NETWORK
TITLE = Station Sicher Pos3.0
      AN    "POS3_0_Prodiag_DB".State.C1;

      =     "HMI_BETR_ART_POS".POS3_0.Status_Sicher;

END_FUNCTION_BLOCK

FUNCTION_BLOCK "Melden_VisuAllgemein"   // FB127, LAD
{ S7_Optimized_Access := 'TRUE' }
// stored: MemoryReserve 100, SetENOAutomatically false
   VAR
      Register_leer : "Teile Status";
      auf_Seite_Richten { S7_SetPoint := 'True'} : Bool;
      Flanke_Bildwechsel { S7_SetPoint := 'True'} : R_TRIG;
      Bild_tmp { S7_SetPoint := 'True'} : DInt;
      WartezeitSicherung_Reset { S7_SetPoint := 'True'} : TON_TIME;
      Flanke_Türe8_schließen { S7_SetPoint := 'True'} : R_TRIG;
      Flanke_Türe8_öffnen { S7_SetPoint := 'True'} : R_TRIG;
   END_VAR
   VAR RETAIN
      Artikelnummer_tmp { ExternalAccessible := 'False'; ExternalVisible := 'False'; ExternalWritable := 'False'} : String;
   END_VAR
   VAR
      VZ_Leerfahren { S7_SetPoint := 'True'} : TON_TIME;
   END_VAR
   VAR_TEMP
      test : Bool;
   END_VAR
BEGIN

REGION Network 1 (SCL): Richten oder Einzelschrittseite aufgerufen
   CASE "HMI_SYS"."Aktueller Bildschirm" OF
       75:
           #auf_Seite_Richten := true;
       ELSE
           #auf_Seite_Richten := false;
   END_CASE;
END_REGION

REGION Network 2 (SCL): Artikel wurde gewechselt


   IF #Artikelnummer_tmp <> "HMI_COM".Artikelnummer_String THEN
       "HMI_COM".Artikel_gewechselt := true;
       #Artikelnummer_tmp := "HMI_COM".Artikelnummer_String;
   ELSIF "HMI_COM".Grundstellung_Gesamt AND  "HMI_COM".Artikel_gewechselt THEN

       "HMI_COM".Artikel_gewechselt := false;

   END_IF;
END_REGION

NETWORK
TITLE = Übergabe Anwahl Richten
      A     #auf_Seite_Richten;
      JC    m003;

      JU    m001;
m003: NOP   0;

      A     "03_Betriebsart_DB"."NOT-HALT OK";
      A     "03_Betriebsart_DB"."Schutztüren OK";
      JCN   m001;


      A     "HMI_COM".Richten_Gesamtanlage;
      JCN   m002;

      SET;
      S     "HMI_BETR_ART_POS".POS3_0.Taster_Anwahl_GS;


m002: NOP   0;

      A     "HMI_BETR_ART_POS".POS3_0.Taster_Anwahl_GS;
      S     "POS3_0_Signal".Station.SK_Freigabe_Richten;
      =     "POS3_0_Signal".Schrittkette.INIT_SQ;
      R     "HMI_BETR_ART_POS".POS3_0.Taster_Anwahl_GS;


      A     "HMI_COM".Richten_Gesamtanlage;
      R     "HMI_COM".Richten_Gesamtanlage;

m001: NOP   0;


NETWORK
TITLE = Tippbetrieb Aktiv
      A     "POS3_0_Signal".Schrittkette.AUTO_ON;


      =     "HMI_COM".Einzelschritt.Status_Anw;


NETWORK
TITLE = Antriebe sind Ein
      SET;

      =     "HMI_COM".Antriebe_sind_EIN;

REGION Network 6 (SCL): Übergabe Türen Not Halt
   // Allgemeine HMI Übergabe 

   "HMI_COM"."NOT-HALT_OK" := "03_Betriebsart_DB"."NOT-HALT OK";
   "HMI_COM".TUERE_OK := "03_Betriebsart_DB"."Schutztüren OK";




   // Übergabe welche Tür ist nicht verriegelt
   REGION Türen


       "HMI_COM".Tür_offen[1] := "DE_Rueckfuehrung_Tuer_1" AND ("03_Betriebsart_DB".BA_Automatik OR "03_Betriebsart_DB".BA_Manuell OR "03_Betriebsart_DB".BA_Richten);
       "HMI_COM".Tür_offen[2] := "DE_Rueckfuehrung_Tuer_2" AND ("03_Betriebsart_DB".BA_Automatik OR "03_Betriebsart_DB".BA_Manuell OR "03_Betriebsart_DB".BA_Richten);
    //   "HMI_COM".Tür_offen[3] := "DE_Rueckfuehrung_Tuer_3" AND ("03_Betriebsart_DB".BA_Automatik OR "03_Betriebsart_DB".BA_Manuell OR "03_Betriebsart_DB".BA_Richten);
    //   "HMI_COM".Tür_offen[4] := "DE_Rueckfuehrung_Tuer_4" AND ("03_Betriebsart_DB".BA_Automatik OR "03_Betriebsart_DB".BA_Manuell OR "03_Betriebsart_DB".BA_Richten);
    //   "HMI_COM".Tür_offen[5] := "DE_Rueckfuehrung_Tuer_5" AND ("03_Betriebsart_DB".BA_Automatik OR "03_Betriebsart_DB".BA_Manuell OR "03_Betriebsart_DB".BA_Richten);
    //   "HMI_COM".Tür_offen[6] := "DE_Rueckfuehrung_Tuer_6" AND ("03_Betriebsart_DB".BA_Automatik OR "03_Betriebsart_DB".BA_Manuell OR "03_Betriebsart_DB".BA_Richten);
    //   "HMI_COM".Tür_offen[7] := "DE2_0_Rückführung Tür 7" AND ("03_Betriebsart_DB".BA_Automatik OR "03_Betriebsart_DB".BA_Manuell OR "03_Betriebsart_DB".BA_Richten);
    //   "HMI_COM".Tür_offen[8] := "DE2_1_Rückführung Tür 8" AND ("03_Betriebsart_DB".BA_Automatik OR "03_Betriebsart_DB".BA_Manuell OR "03_Betriebsart_DB".BA_Richten);
    (*   "HMI_COM".Tür_offen[9] := "DE2_1_Rückführung Tür 8" AND ("03_Betriebsart_DB".BA_Automatik OR "03_Betriebsart_DB".BA_Manuell OR "03_Betriebsart_DB".BA_Richten);
       "HMI_COM".Tür_offen[10] := "DE2_1_Rückführung Tür 8" AND ("03_Betriebsart_DB".BA_Automatik OR "03_Betriebsart_DB".BA_Manuell OR "03_Betriebsart_DB".BA_Richten);
       "HMI_COM".Tür_offen[11] := "DE2_1_Rückführung Tür 8" AND ("03_Betriebsart_DB".BA_Automatik OR "03_Betriebsart_DB".BA_Manuell OR "03_Betriebsart_DB".BA_Richten);
       "HMI_COM".Tür_offen[12] := "DE2_1_Rückführung Tür 8" AND ("03_Betriebsart_DB".BA_Automatik OR "03_Betriebsart_DB".BA_Manuell OR "03_Betriebsart_DB".BA_Richten);
       "HMI_COM".Tür_offen[13] := "DE2_1_Rückführung Tür 8" AND ("03_Betriebsart_DB".BA_Automatik OR "03_Betriebsart_DB".BA_Manuell OR "03_Betriebsart_DB".BA_Richten);
       "HMI_COM".Tür_offen[14] := "DE2_1_Rückführung Tür 8" AND ("03_Betriebsart_DB".BA_Automatik OR "03_Betriebsart_DB".BA_Manuell OR "03_Betriebsart_DB".BA_Richten);
       "HMI_COM".Tür_offen[15] := "DE2_1_Rückführung Tür 8" AND ("03_Betriebsart_DB".BA_Automatik OR "03_Betriebsart_DB".BA_Manuell OR "03_Betriebsart_DB".BA_Richten); *)
    //   "HMI_COM".Tür_offen[16] := "DE2_1_Rückführung Tür 8" AND ("03_Betriebsart_DB".BA_Automatik OR "03_Betriebsart_DB".BA_Manuell OR "03_Betriebsart_DB".BA_Richten);

   END_REGION
END_REGION

REGION Network 7 (SCL): Rücksetzen der Stationen bei Grundbild



   #Flanke_Bildwechsel(CLK:="03_Betriebsart_DB".BA_Manuell AND #Bild_tmp <> "HMI_SYS"."Aktueller Bildschirm" );



   IF #Flanke_Bildwechsel.Q THEN

       #Bild_tmp := "HMI_SYS"."Aktueller Bildschirm";

    //IF ("HMI_SYS"."Aktueller Bildschirm" = 10125) OR ("03_Betriebsart_DB"."NOT-HALT OK" = false) THEN

       "HMI_COM".Manuell_Zylinder1.Status := 0;
       "HMI_COM".Manuell_Zylinder2.Status := 0;
       "HMI_COM".Manuell_Zylinder3.Status := 0;
       "HMI_COM".Manuell_Zylinder4.Status := 0;

       "HMI_COM".Manuell_Zylinder1.GS := FALSE;
       "HMI_COM".Manuell_Zylinder1.AS1 := FALSE;
       "HMI_COM".Manuell_Zylinder2.GS := FALSE;
       "HMI_COM".Manuell_Zylinder2.AS1 := FALSE;
       "HMI_COM".Manuell_Zylinder3.GS := FALSE;
       "HMI_COM".Manuell_Zylinder3.AS1 := FALSE;
       "HMI_COM".Manuell_Zylinder4.GS := FALSE;
       "HMI_COM".Manuell_Zylinder4.AS1 := FALSE;

      "HMI_COM".Manuell_Zylinder1.DA_GS := FALSE;
       "HMI_COM".Manuell_Zylinder1.DA_AS1 := FALSE;
       "HMI_COM".Manuell_Zylinder2.DA_GS := FALSE;
       "HMI_COM".Manuell_Zylinder2.DA_AS1 := FALSE;
       "HMI_COM".Manuell_Zylinder3.DA_GS := FALSE;
       "HMI_COM".Manuell_Zylinder3.DA_AS1 := FALSE;
       "HMI_COM".Manuell_Zylinder4.DA_GS := FALSE;
       "HMI_COM".Manuell_Zylinder4.DA_AS1 := FALSE;
     END_IF;
END_REGION

REGION Network 8 (SCL): Übertragung und Verwaltung Register



   "HMI_COM".Speichern_Register := false;
END_REGION

REGION Network 9 (SCL): Rucksetzen wenn Register nicht gelöscht
   IF (("HMI_SYS"."Aktueller Bildschirm" = 10001) OR ("HMI_SYS"."Aktueller Bildschirm" = 10010) OR ("HMI_SYS"."Aktueller Bildschirm" = 10020)
       OR ("HMI_SYS"."Aktueller Bildschirm" = 10030)) THEN

       "HMI_BETR_ART_POS".POS3_0.Taster_Reset_Teilestatus := FALSE;
       "HMI_BETR_ART_POS".POS3_1.Taster_Reset_Teilestatus := FALSE;
       "HMI_BETR_ART_POS".POS3_2.Taster_Reset_Teilestatus := FALSE;
       "HMI_BETR_ART_POS".POS3_3.Taster_Reset_Teilestatus := FALSE;
       "HMI_BETR_ART_POS".POS3_4.Taster_Reset_Teilestatus := FALSE;
       "HMI_BETR_ART_POS".POS4_0_Zuführung.Taster_Reset_Teilestatus := FALSE;
       "HMI_BETR_ART_POS".POS5_0_Zuführung.Taster_Reset_Teilestatus := FALSE;
       "HMI_BETR_ART_POS".POS5_0.Taster_Reset_Teilestatus := FALSE;
       "HMI_BETR_ART_POS".POS6_0.Taster_Reset_Teilestatus := FALSE;
       "HMI_BETR_ART_POS".POS7_0.Taster_Reset_Teilestatus := FALSE;
       "HMI_BETR_ART_POS".POS7_1.Taster_Reset_Teilestatus := FALSE;
       "HMI_BETR_ART_POS".POS7_2.Taster_Reset_Teilestatus := FALSE;
       "HMI_BETR_ART_POS".POS7_3.Taster_Reset_Teilestatus := FALSE;
       "HMI_BETR_ART_POS".POS7_4.Taster_Reset_Teilestatus := FALSE;
       "HMI_BETR_ART_POS".POS8_0.Taster_Reset_Teilestatus := FALSE;
       "HMI_BETR_ART_POS".POS9_0.Taster_Reset_Teilestatus := FALSE;
       "HMI_BETR_ART_POS".POS9_1.Taster_Reset_Teilestatus := FALSE;
       "HMI_BETR_ART_POS".POS9_2.Taster_Reset_Teilestatus := FALSE;
       "HMI_BETR_ART_POS".POS9_3.Taster_Reset_Teilestatus := FALSE;
       "HMI_BETR_ART_POS".POS9_4.Taster_Reset_Teilestatus := FALSE;
       "HMI_BETR_ART_POS".POS9_5.Taster_Reset_Teilestatus := FALSE;
       "HMI_BETR_ART_POS".POS9_6.Taster_Reset_Teilestatus := FALSE;
       "HMI_BETR_ART_POS".POS10_0.Taster_Reset_Teilestatus := FALSE;
       "HMI_BETR_ART_POS".POS11.Taster_Reset_Teilestatus := FALSE;
       "HMI_BETR_ART_POS".POS12.Taster_Reset_Teilestatus := FALSE;

   END_IF;
END_REGION

REGION Network 10 (SCL): Leerfahren
   "HMI_Signale".Leerfahren_angewaehlt := "HMI_COM".Leerfahren_angewaehlt;

   #VZ_Leerfahren(IN := "HMI_COM".Leerfahren_ende,
                  PT := t#3s);

   IF #VZ_Leerfahren.Q OR "HMI_COM".Leerfahren_angewaehlt = false THEN

       "HMI_COM".Leerfahren_ende := FALSE;
       "HMI_Signale".Leerfahren_ende := false;
       "HMI_COM".Leerfahren_angewaehlt := false;

       "HMI_COM".Leerfahren_laeuft := false; 
       "POS3_0_Signal".Station.SK_Freigabe_Auto := false;




   END_IF;
END_REGION

REGION Network 11 (SCL): Bildaufrufe


       // Bei Not-Aus Aufruf Grundbild
       IF "03_Betriebsart_DB".BA_0_FP = TRUE OR
           "03_Betriebsart_DB"."NOT-HALT_FN" = TRUE OR
           "03_Betriebsart_DB".Schutztüren_FN = TRUE THEN
           "HMI_SYS".Screen_Name := WSTRING#'B10001_Hauptbild';
       END_IF;


       // Bei BA Manuell Auswahlbild aufrufen
       IF "03_Betriebsart_DB".BA_Manuell_FP = TRUE THEN
           "HMI_SYS".Screen_Name := WSTRING#'B10020_Manuell Auswahl';
       END_IF;


       // Bei BA Richten Auswahlbild aufrufen
       IF "03_Betriebsart_DB".BA_Richten_FP = TRUE THEN
           "HMI_SYS".Screen_Name := WSTRING#'B10075_Übersicht Richten Stationen';
       END_IF;


       // Bei BA Automatik Auswahlbild aufrufen
       IF "03_Betriebsart_DB".BA_Automatik_FP = TRUE THEN
           "HMI_SYS".Screen_Name := WSTRING#'B10010_Automatik';
       END_IF;


       // Bei BA Verwaltung Auswahlbild aufrufen
       IF "03_Betriebsart_DB".BA_Verwaltung_FP = TRUE THEN
           "HMI_SYS".Screen_Name := WSTRING#'B10030_Übersicht Verwaltung';
       END_IF;
END_REGION

REGION Network 12 (SCL): DE +HS1=AN-22T1 Selektivmodul
   #test := NOT "DE_Selektivmodul_OK";

   #WartezeitSicherung_Reset(IN:=#test,
                             PT:=t#25s);





   IF #WartezeitSicherung_Reset.Q = False AND "DE_Selektivmodul_OK"= false THEN
       "HMI_COM".Status_24V_Sicherung := 3;
   ELSIF "DE_Selektivmodul_OK" = false AND "HMI_COM".Status_24V_Sicherung <> 2 THEN
       "HMI_COM".Status_24V_Sicherung  := 0;
   ELSIF "DE_Selektivmodul_OK" = false AND "HMI_COM".Status_24V_Sicherung = 2 THEN
       "DA_Selektivmodul Reset" := true;
   ELSIF "DE_Selektivmodul_OK" THEN
       "HMI_COM".Status_24V_Sicherung := 1;
       "DA_Selektivmodul Reset" := false;
   END_IF;
END_REGION

REGION Network 13 (SCL): nur zum testen
   (* IF "HMI_COM".HMI_Achse_Steuerung.E_jog_pos THEN

       "Pos3_0_Signal".Y_Achse_1.E_jog_pos := true;
       "Pos3_0_Signal".Y_Achse_2.E_jog_pos := true;
       "Pos3_0_Signal".Y_Achse_3.E_jog_pos := true;
       "Pos3_0_Signal".Y_Achse_4.E_jog_pos := true;
       "Pos3_0_Signal".Y_Achse_1.E_jog_neg := 0;
       "Pos3_0_Signal".Y_Achse_2.E_jog_neg := 0;
       "Pos3_0_Signal".Y_Achse_3.E_jog_neg := 0;
       "Pos3_0_Signal".Y_Achse_4.E_jog_neg := 0;

   ELSIF "HMI_COM".HMI_Achse_Steuerung.E_jog_neg THEN


       "Pos3_0_Signal".Y_Achse_1.E_jog_neg := true;
       "Pos3_0_Signal".Y_Achse_2.E_jog_neg := true;
       "Pos3_0_Signal".Y_Achse_3.E_jog_neg := true;
       "Pos3_0_Signal".Y_Achse_4.E_jog_neg := true;

       "Pos3_0_Signal".Y_Achse_1.E_jog_pos := 0;
       "Pos3_0_Signal".Y_Achse_2.E_jog_pos := 0;
       "Pos3_0_Signal".Y_Achse_3.E_jog_pos := 0;
       "Pos3_0_Signal".Y_Achse_4.E_jog_pos := 0;

   ELSE
       "Pos3_0_Signal".Y_Achse_1.E_jog_neg := 0;
       "Pos3_0_Signal".Y_Achse_2.E_jog_neg := 0;
       "Pos3_0_Signal".Y_Achse_3.E_jog_neg := 0;
       "Pos3_0_Signal".Y_Achse_4.E_jog_neg := 0;
       "Pos3_0_Signal".Y_Achse_1.E_jog_pos := 0;
       "Pos3_0_Signal".Y_Achse_2.E_jog_pos := 0;
       "Pos3_0_Signal".Y_Achse_3.E_jog_pos := 0;
       "Pos3_0_Signal".Y_Achse_4.E_jog_pos := 0;
   END_IF; *)

   // "HMI_COM".Manuell_Zylinder1.GS := false;
   // "HMI_COM".Manuell_Zylinder1.AS1 := false;
   // "HMI_COM".Manuell_Zylinder2.GS := false;
   // "HMI_COM".Manuell_Zylinder2.AS1 := false;
   // "HMI_COM".Manuell_Zylinder3.GS := false;
   // "HMI_COM".Manuell_Zylinder3.AS1 := false;
   // "HMI_COM".Manuell_Zylinder4.GS := false;
   // "HMI_COM".Manuell_Zylinder4.AS1 := false;
END_REGION

REGION Network 14 (SCL): Übergabe Taktzeiten Stationen
   "HMI_COM".Taktzeit[0] := "POS3_0_Signal".Taktzeit[0];
END_REGION

REGION Network 15 (SCL): Rücksetzten Messmittelabläufe
   IF ("HMI_COM".Abläufe_Messmittel < 1) OR "03_Betriebsart_DB".Stopp_Taste = false THEN
       "HMI_COM".Messmittel_ein := false;
       ;
   END_IF;


   IF ("HMI_COM".Abläufe_Messmittel_Rundlauf < 1) OR "03_Betriebsart_DB".Stopp_Taste = false THEN
       "HMI_COM".Messmittel_Rundlauf_ein := false;
       ;
   END_IF;
END_REGION
END_FUNCTION_BLOCK

FUNCTION "Störmeldungen" : Void   // FC512, STL
TITLE = Störmeldungen
{ S7_Optimized_Access := 'FALSE' }
// Störmeldungsbaustein: Hier befinden sich alle Störungen zusammengefasst zur 
// Sammelstörung und alle Störungen, die nicht in FB`s aufgelistet wurden.
// stored: AutoNumber false
   VAR_TEMP
      retval : Int;
      keine_Störung : Bool;
   END_VAR
BEGIN

NETWORK
TITLE = Sammelstörung Anlage
      A     "ProDiag_Allgemein_DB".State.C1;
      O     "POS3_0_Prodiag_DB".State.C1;



// Schrittketten in Störung (Interlock oder Supervision)
      O     "POS3_0_Signal".Schrittkette.ERR_FLT;

      =     "HMI_Signale".Sammelstoerung;


NETWORK
TITLE = Stop von Störmeldungen



      CLR;
      S     "HMI_Signale".Stop_Von_Stoermeldung;

      A     "03_Betriebsart_DB".ACK_Taste;
      R     "HMI_Signale".Stop_Von_Stoermeldung;
END_FUNCTION

FUNCTION_BLOCK "Leuchtmelder Ampel"
{ S7_Optimized_Access := 'TRUE' }
VERSION : 0.1
   VAR 
      Ampelbaustein_MG_Instance : "Ampelbaustein_MG";
      OUT_Ampel_rot { S7_SetPoint := 'True'} : Bool;
      OUT_Ampel_gelb { S7_SetPoint := 'True'} : Bool;
      OUT_Ampel_gruen { S7_SetPoint := 'True'} : Bool;
      OUT_Akkustik { S7_SetPoint := 'True'} : Bool;
   END_VAR

   VAR_TEMP 
      TEMP_IO_Kiste_Voll : Bool;
   END_VAR


BEGIN
	// Anlagenbeleuchtung 
	"DA_Anlagenbeleuchtung" :=  "HMI_COM".Anlagenbeleuchtung_EIN ;
	
	
	// Ampel
	// 
	
	
	    #TEMP_IO_Kiste_Voll := FALSE;
	
	
	    #Ampelbaustein_MG_Instance(Sammelstoerung:="HMI_Signale".Sammelstoerung,
	                               BA_0:="03_Betriebsart_DB".BA_0,
	                               BA_A:="03_Betriebsart_DB".BA_Automatik,
	                               BA_M:="03_Betriebsart_DB".BA_Manuell,
	                               BA_R:="03_Betriebsart_DB".BA_Richten,
	                               BA_V:="03_Betriebsart_DB".BA_Verwaltung,
	                               Ablauf_ist_aktiv:="HMI_Signale".Freigabe_Zyklus,
	                               Blinker:="Clock_1Hz",
	                               Ampel_rot=> #OUT_Ampel_rot,
	                               Ampel_gelb=> #OUT_Ampel_gelb,
	                               Ampel_gruen=> #OUT_Ampel_gruen,
	                               Akkustik=> #OUT_Akkustik);
	//        Trigger 1   Trigger 2
	// AUS    LO          LO
	// ROT    HI          LO
	// GELB   HI          HI
	// GRÜN   LO          HI
	// 
	    IF #OUT_Ampel_rot AND
	        "03_Betriebsart_DB".BA_0 = false THEN
	        "DA_Anlagenzustand_Trigger_1" := true;
	        "DA_Anlagenzustand_Trigger_2" := false;
	    ELSIF #OUT_Ampel_gelb AND
	        "03_Betriebsart_DB".BA_0 = false THEN
	        "DA_Anlagenzustand_Trigger_1" := true;
	        "DA_Anlagenzustand_Trigger_2" := true;
	    ELSIF #OUT_Ampel_gruen AND
	        "03_Betriebsart_DB".BA_0 = false THEN
	        "DA_Anlagenzustand_Trigger_1" := false;
	        "DA_Anlagenzustand_Trigger_2" := true;
	    ELSE
	        "DA_Anlagenzustand_Trigger_1" := false;
	        "DA_Anlagenzustand_Trigger_2" := false;
	    END_IF;
END_FUNCTION_BLOCK

FUNCTION_BLOCK "Ampelbaustein_MG"   // FB145, STL
{ S7_Optimized_Access := 'FALSE' }
// stored: AutoNumber false
   VAR_INPUT
      Sammelstoerung : Bool;
      BA_0 : Bool;
      BA_A : Bool;
      BA_M : Bool;
      BA_R : Bool;
      BA_V : Bool;
      Ablauf_ist_aktiv : Bool;
      Blinker : Bool;
   END_VAR
   VAR_OUTPUT
      Ampel_rot : Bool;
      Ampel_gelb : Bool;
      Ampel_gruen : Bool;
      Akkustik : Bool;
   END_VAR
   VAR
      Timer_Hupe_EIN { S7_SetPoint := 'True'} : TON_TIME;
      Timer_Hupe_Aus { S7_SetPoint := 'True'} : TON_TIME;
      Ampel_Zustand : Int;
   END_VAR
BEGIN

NETWORK
TITLE = Ampel Betriebsart 0-4
      L     0;
      T     #Ampel_Zustand;

// Grün
      A     #Ablauf_ist_aktiv;
      A     #BA_A;
      AN    #Sammelstoerung;
      JCN   zustand_rot;
      L     1;
      T     #Ampel_Zustand;
      JU    auswertung;

// Rot
zustand_rot:NOP   0;
      A     #Sammelstoerung;
      JCN   zustand_gelb;
      L     2;
      T     #Ampel_Zustand;
      JU    auswertung;


// Gelb
zustand_gelb:NOP   0;
      A     #BA_A;
      O     #BA_M;
      O     #BA_V;
      O     #BA_R;
      JCN   auswertung;
      L     3;
      T     #Ampel_Zustand;

// Aus
zustand_Aus:NOP   0;
      A     #BA_0;
      JCN   auswertung;
      L     4;
      T     #Ampel_Zustand;





NETWORK
TITLE = Sprungliste in die jewilige Ampelbeschaltung (wie case anweisung)
auswertung:NOP   0;
      L     #Ampel_Zustand;
      JL    end;
      JU    NOP;
      JU    grün;
      JU    rot;
      JU    gelb;
      JU    Aus;
end:  JU    ENDE;

NETWORK
TITLE = Nicht definiert
NOP:  NOP   0;


      CLR;
      =     #Ampel_gelb;
      =     #Ampel_rot;
      =     #Ampel_gruen;
      =     #Akkustik;



      JU    ENDE;


NETWORK
TITLE = Grün
grün: NOP   0;
      SET;
      =     #Ampel_gruen;
      CLR;
      =     #Ampel_gelb;
      =     #Ampel_rot;
      =     #Akkustik;
      JU    ENDE;


NETWORK
TITLE = Rot
rot:  NOP   0;
      SET;
      =     #Ampel_rot;
      CLR;
      =     #Ampel_gelb;
      =     #Ampel_gruen;
      =     #Akkustik;
      JU    ENDE;

NETWORK
TITLE = Gelb
gelb: NOP   0;
      SET;
      =     #Ampel_gelb;
      CLR;
      =     #Ampel_rot;
      =     #Ampel_gruen;
      =     #Akkustik;

      JU    ENDE;

NETWORK
TITLE = Aus
Aus:  NOP   0;
      SET;

      CLR;
      =     #Ampel_rot;
      =     #Ampel_gelb;
      =     #Ampel_gruen;
      =     #Akkustik;

      JU    ENDE;

NETWORK
TITLE = ENDE Sprungleiste
ENDE: NOP   0;


NETWORK
TITLE = Störungshupe
      CALL  #Timer_Hupe_EIN
      ( IN := #Sammelstoerung,
        PT := T#5M,
        Q  := ,
        ET := 
      );

      CALL  #Timer_Hupe_Aus
      ( IN := #Sammelstoerung,
        PT := T#10M,
        Q  := ,
        ET := 
      );

      A     #Sammelstoerung;
      A     #Blinker;
//      U     #Timer_Hupe_EIN.Q
//      UN    #Timer_Hupe_Aus.Q
      A     #BA_A;
      =     #Akkustik;

END_FUNCTION_BLOCK

FUNCTION_BLOCK "FB002_LabView"
{ S7_Optimized_Access := 'TRUE' }
VERSION : 0.1

BEGIN
	
	// Lebenszeichen 
	IF "FL_Clock_1Hz"  THEN
	    "DB020_Com LabView".A_Lebenszeichen := "DB020_Com LabView".A_Lebenszeichen + 1;
	    IF "DB020_Com LabView".A_Lebenszeichen > 9999 THEN
	        "DB020_Com LabView".A_Lebenszeichen := 1;
	    END_IF;
	END_IF;
	
	// Betriebsart
	
	"DB020_Com LabView".A_Betriebsart := "03_Betriebsart_DB".Betriebsart;
	
	
	// Wenn Messung fertig, Signal "Messung läuft" zurücksetzen
	IF "DB020_Com LabView"."E_Messgerät ist bereit und verbunden" THEN
	    "DB020_Com LabView".E_4_4 := false;
	END_IF;
	 
	
	"DB020_Com LabView".A_Steckzyklen_Soll := "POS3_0_Signal".Sollzyklen;
	"DB020_Com LabView".A_Steckzyklen_Ist := "POS3_0_Signal".Istzyklen;
	
	"DB020_Com LabView".A_Achse_Istposition := "POS3_0_Signal"."-1001T1 Oriental_Steuerung".A_FBposition;
	"DB020_Com LabView".A_Achse_Drehmoment :=  "POS3_0_Signal"."-1001T1 Oriental_Steuerung".A_TorqueMonitor;
	
	
	"DB020_Com LabView".A_Drehachse_Istposition  := "POS3_0_Signal"."-1002T1 Oriental_Steuerung".A_FBposition;
	"DB020_Com LabView".A_Drehachse_Drehmoment :=  "POS3_0_Signal"."-1002T1 Oriental_Steuerung".A_TorqueMonitor;
	
	"DB020_Com LabView".A_Wegmessung_Ausgleichszylinder_Istwert := "POS3_0_Signal"."-POS3.0_Wegmessung_Ausgleichszylinder_Istwert_Rohwert";
	
	"DB020_Com LabView".A_Kraftsensor_Istwert := "POS3_0_Signal"."-1012B1 Kraftsensor";
	
	
	"DB020_Com LabView".A_Regelventil_Ausgleichszylinder_Istwert := "POS3_0_Signal"."-POS3_0_Regelventil_Ausgleichszylinder_Istwert";
	
	"DB020_Com LabView".A_Regelventil_Überlastzylinder_Istwert := "POS3_0_Signal"."-POS3_0_Regelventil_Überlastzylinder_Istwert";
	
	 
END_FUNCTION_BLOCK

FUNCTION_BLOCK "Verwaltung_Teiledaten_FB"
{ S7_Optimized_Access := 'TRUE' }
VERSION : 0.1

BEGIN
	IF "Verwaltung_Teiledaten"."Taster Achse Position GS übernehmen" THEN
	    "Verwaltung_Teiledaten"."Achse Position GS" := "POS3_0_Signal"."-1001T1 Oriental_Steuerung".A_FBposition;
	    "Verwaltung_Teiledaten"."Taster Achse Position GS übernehmen" := false;
	END_IF;
	
	
	IF "Verwaltung_Teiledaten"."Taster Achse Position AS übernehmen" THEN
	    "Verwaltung_Teiledaten"."Achse Position AS" := "POS3_0_Signal"."-1001T1 Oriental_Steuerung".A_FBposition;
	    "Verwaltung_Teiledaten"."Taster Achse Position AS übernehmen" := false;
	END_IF;
	
	
	IF "Verwaltung_Teiledaten"."Taster Drehantrieb Position GS übernehmen" THEN
	    "Verwaltung_Teiledaten"."Drehantrieb Position GS" := 0.0;
	    "POS3_0_Signal"."-1002T1 Oriental_E_P-Preset" := true;
	    "Verwaltung_Teiledaten"."Taster Drehantrieb Position GS übernehmen" := false;
	END_IF;
	
	
	
	IF "Verwaltung_Teiledaten"."Taster Drehantrieb Position AS1 übernehmen" THEN
	    "Verwaltung_Teiledaten"."Drehantrieb Position AS1" := "POS3_0_Signal"."-1002T1 Oriental_Absolute_Position";
	    "Verwaltung_Teiledaten"."Taster Drehantrieb Position AS1 übernehmen" := false;
	END_IF;
	
	
	IF "Verwaltung_Teiledaten"."Taster Drehantrieb Position AS2 übernehmen" THEN
	    "Verwaltung_Teiledaten"."Drehantrieb Position AS2" := "POS3_0_Signal"."-1002T1 Oriental_Absolute_Position";
	    "Verwaltung_Teiledaten"."Taster Drehantrieb Position AS2 übernehmen" := false;
	END_IF;
	
	
	IF "Verwaltung_Teiledaten"."Taster Wegmessung Ausgleichszylinder Position AS1 übernehmen" THEN
	    "Verwaltung_Teiledaten"."Wegmessung_Ausgleichszylinder maximale Abweichung GS" := "POS3_0_Signal"."-POS3.0_Wegmessung_Ausgleichszylinder_Istwert_Rohwert";
	    "Verwaltung_Teiledaten"."Taster Wegmessung Ausgleichszylinder Position AS1 übernehmen" := false;
	END_IF;
	
	
	"POS3_0_Signal"."Wartezeit Soll gesteckt" := DINT_TO_TIME(REAL_TO_DINT("Verwaltung_Teiledaten"."Wartezeit gesteckt" * 1000.0));
	
	
END_FUNCTION_BLOCK

FUNCTION_BLOCK "01_Alle_Zaehler"   // FB48, FBD
{ S7_Optimized_Access := 'TRUE' }
// stored: MemoryReserve 100, SetENOAutomatically false
   VAR
      Zaehlsignal_Gesamt : Bool;
      Zaehlsignal_IO : Bool;
      Zaehlsignal_NIO : Bool;
      Zaehlsignal_NIO_LabView : Bool;
      "Zaehlsignal_IO_1 Palette 1" : Bool;
      "Zaehlsignal_IO_2 Palette 2" : Bool;
      "Zaehlsignal_IO_3 Palette 3" : Bool;
      "Zaehlsignal_IO_4 Palette 4" : Bool;
      "Zaehlsignal_IO_5 Palette 5" : Bool;
      "Zaehlsignal_NIO_1_Palette NIO" : Bool;
      Zaehlsignal_NIO_2 : Bool;
      Zaehlsignal_NIO_3 : Bool;
      Zaehlsignal_NIO_4 : Bool;
      Zaehlsignal_NIO_5 : Bool;
      Zaehlsignal_NIO_6 : Bool;
   END_VAR
BEGIN

NETWORK
TITLE = Zählerstand Teile Gesamt
      CALL  "Zählerfunktion >1000"
      ( Schichtzaehler_Reset  := "HMI_COM".Reset_Schichtzaehler,
        Auftragszaehler_Reset := "HMI_COM".Reset_Auftragszaehler,
        Schichtzaehler        := "HMI_Statistik"."Zaehler Alle Teile".Schichtzaehler,
        Auftragszaehler       := "HMI_Statistik"."Zaehler Alle Teile".Auftragszaehler,
        Gesamtzaehler         := "HMI_Statistik"."Zaehler Alle Teile".Gesamtzaehler,
        Zaehlsignal           := #Zaehlsignal_Gesamt
      );



NETWORK
TITLE = Zählerstand IO gesamt
      CALL  "Zählerfunktion >1000"
      ( Schichtzaehler_Reset  := "HMI_COM".Reset_Schichtzaehler,
        Auftragszaehler_Reset := "HMI_COM".Reset_Auftragszaehler,
        Schichtzaehler        := "HMI_Statistik"."Zaehler IO Teile".Schichtzaehler,
        Auftragszaehler       := "HMI_Statistik"."Zaehler IO Teile".Auftragszaehler,
        Gesamtzaehler         := "HMI_Statistik"."Zaehler IO Teile".Gesamtzaehler,
        Zaehlsignal           := #Zaehlsignal_IO
      );



NETWORK
TITLE = Zählerstand NIO gesamt

      CALL  "Zählerfunktion >1000"
      ( Schichtzaehler_Reset  := "HMI_COM".Reset_Schichtzaehler,
        Auftragszaehler_Reset := "HMI_COM".Reset_Auftragszaehler,
        Schichtzaehler        := "HMI_Statistik"."Zaehler NIO Teile".Schichtzaehler,
        Auftragszaehler       := "HMI_Statistik"."Zaehler NIO Teile".Auftragszaehler,
        Gesamtzaehler         := "HMI_Statistik"."Zaehler NIO Teile".Gesamtzaehler,
        Zaehlsignal           := #Zaehlsignal_NIO
      );



NETWORK
TITLE = IO Zähler 1

      CALL  "Zählerfunktion >1000"
      ( Schichtzaehler_Reset  := "HMI_COM".Reset_Schichtzaehler,
        Auftragszaehler_Reset := "HMI_COM".Reset_Auftragszaehler,
        Schichtzaehler        := "HMI_Statistik"."IO 1".Schichtzaehler,
        Auftragszaehler       := "HMI_Statistik"."IO 1".Auftragszaehler,
        Gesamtzaehler         := "HMI_Statistik"."IO 1".Gesamtzaehler,
        Zaehlsignal           := #"Zaehlsignal_IO_1 Palette 1"
      );


NETWORK
TITLE = IO Zähler 2

      CALL  "Zählerfunktion >1000"
      ( Schichtzaehler_Reset  := "HMI_COM".Reset_Schichtzaehler,
        Auftragszaehler_Reset := "HMI_COM".Reset_Auftragszaehler,
        Schichtzaehler        := "HMI_Statistik"."IO 2".Schichtzaehler,
        Auftragszaehler       := "HMI_Statistik"."IO 2".Auftragszaehler,
        Gesamtzaehler         := "HMI_Statistik"."IO 2".Gesamtzaehler,
        Zaehlsignal           := #"Zaehlsignal_IO_2 Palette 2"
      );




NETWORK
TITLE = IO Zähler 3

      CALL  "Zählerfunktion >1000"
      ( Schichtzaehler_Reset  := "HMI_COM".Reset_Schichtzaehler,
        Auftragszaehler_Reset := "HMI_COM".Reset_Auftragszaehler,
        Schichtzaehler        := "HMI_Statistik"."IO 3".Schichtzaehler,
        Auftragszaehler       := "HMI_Statistik"."IO 3".Auftragszaehler,
        Gesamtzaehler         := "HMI_Statistik"."IO 3".Gesamtzaehler,
        Zaehlsignal           := #"Zaehlsignal_IO_3 Palette 3"
      );




NETWORK
TITLE = IO Zähler 4

      CALL  "Zählerfunktion >1000"
      ( Schichtzaehler_Reset  := "HMI_COM".Reset_Schichtzaehler,
        Auftragszaehler_Reset := "HMI_COM".Reset_Auftragszaehler,
        Schichtzaehler        := "HMI_Statistik"."IO 4".Schichtzaehler,
        Auftragszaehler       := "HMI_Statistik"."IO 4".Auftragszaehler,
        Gesamtzaehler         := "HMI_Statistik"."IO 4".Gesamtzaehler,
        Zaehlsignal           := #"Zaehlsignal_IO_4 Palette 4"
      );




NETWORK
TITLE = IO Zähler 5

      CALL  "Zählerfunktion >1000"
      ( Schichtzaehler_Reset  := "HMI_COM".Reset_Schichtzaehler,
        Auftragszaehler_Reset := "HMI_COM".Reset_Auftragszaehler,
        Schichtzaehler        := "HMI_Statistik"."IO 5".Schichtzaehler,
        Auftragszaehler       := "HMI_Statistik"."IO 5".Auftragszaehler,
        Gesamtzaehler         := "HMI_Statistik"."IO 5".Gesamtzaehler,
        Zaehlsignal           := #"Zaehlsignal_IO_5 Palette 5"
      );




NETWORK
TITLE = NIO Zähler 1

      CALL  "Zählerfunktion >1000"
      ( Schichtzaehler_Reset  := "HMI_COM".Reset_Schichtzaehler,
        Auftragszaehler_Reset := "HMI_COM".Reset_Auftragszaehler,
        Schichtzaehler        := "HMI_Statistik"."NIO 1".Schichtzaehler,
        Auftragszaehler       := "HMI_Statistik"."NIO 1".Auftragszaehler,
        Gesamtzaehler         := "HMI_Statistik"."NIO 1".Gesamtzaehler,
        Zaehlsignal           := #"Zaehlsignal_NIO_1_Palette NIO"
      );


NETWORK
TITLE = NIO Zähler 2

      CALL  "Zählerfunktion >1000"
      ( Schichtzaehler_Reset  := "HMI_COM".Reset_Schichtzaehler,
        Auftragszaehler_Reset := "HMI_COM".Reset_Auftragszaehler,
        Schichtzaehler        := "HMI_Statistik"."NIO 2".Schichtzaehler,
        Auftragszaehler       := "HMI_Statistik"."NIO 2".Auftragszaehler,
        Gesamtzaehler         := "HMI_Statistik"."NIO 2".Gesamtzaehler,
        Zaehlsignal           := #Zaehlsignal_NIO_2
      );


NETWORK
TITLE = NIO Zähler 3

      CALL  "Zählerfunktion >1000"
      ( Schichtzaehler_Reset  := "HMI_COM".Reset_Schichtzaehler,
        Auftragszaehler_Reset := "HMI_COM".Reset_Auftragszaehler,
        Schichtzaehler        := "HMI_Statistik"."NIO 3".Schichtzaehler,
        Auftragszaehler       := "HMI_Statistik"."NIO 3".Auftragszaehler,
        Gesamtzaehler         := "HMI_Statistik"."NIO 3".Gesamtzaehler,
        Zaehlsignal           := #Zaehlsignal_NIO_3
      );


NETWORK
TITLE = NIO Zähler 4

      CALL  "Zählerfunktion >1000"
      ( Schichtzaehler_Reset  := "HMI_COM".Reset_Schichtzaehler,
        Auftragszaehler_Reset := "HMI_COM".Reset_Auftragszaehler,
        Schichtzaehler        := "HMI_Statistik"."NIO 4".Schichtzaehler,
        Auftragszaehler       := "HMI_Statistik"."NIO 4".Auftragszaehler,
        Gesamtzaehler         := "HMI_Statistik"."NIO 4".Gesamtzaehler,
        Zaehlsignal           := #Zaehlsignal_NIO_4
      );




NETWORK
TITLE = NIO Zähler 5

      CALL  "Zählerfunktion >1000"
      ( Schichtzaehler_Reset  := "HMI_COM".Reset_Schichtzaehler,
        Auftragszaehler_Reset := "HMI_COM".Reset_Auftragszaehler,
        Schichtzaehler        := "HMI_Statistik"."NIO 5".Schichtzaehler,
        Auftragszaehler       := "HMI_Statistik"."NIO 5".Auftragszaehler,
        Gesamtzaehler         := "HMI_Statistik"."NIO 5".Gesamtzaehler,
        Zaehlsignal           := #Zaehlsignal_NIO_5
      );


REGION Network 14 (SCL): Reset Taster
   IF "HMI_COM".Reset_Schichtzaehler THEN
       "HMI_COM".Reset_Schichtzaehler := false;
   END_IF;

   IF "HMI_COM".Reset_Auftragszaehler THEN
       "HMI_COM".Reset_Auftragszaehler := false;
   END_IF;
END_REGION
END_FUNCTION_BLOCK

FUNCTION_BLOCK "02_Wartungszaehler"
TITLE = Wartungszähler
{ S7_Optimized_Access := 'TRUE' }
AUTHOR : Falter
FAMILY : HMI
VERSION : 1.0
//Zählerbaustein für Anlgenwartung 25.01.2024
   VAR 
      Wartungszähler_Positionierachse_Zyklen { S7_SetPoint := 'False'} : "FB_Wartungszähler_Zyklen";
      Wartungszähler_Drehachse_Zyklen { S7_SetPoint := 'False'} : "FB_Wartungszähler_Zyklen";
      Wartungszähler_Positionierachse_Weg { S7_SetPoint := 'False'} : "FB_Wartungszähler_Weg";
      Wartungszähler_Drehachse_Weg { S7_SetPoint := 'False'} : "FB_Wartungszähler_Weg";
   END_VAR
   VAR RETAIN
      Positionierachse_Weg { S7_SetPoint := 'True'} : DInt;
      Drehachse_Weg { S7_SetPoint := 'True'} : DInt;
   END_VAR


BEGIN
	
	
	REGION Positionierachse Zyklen
	     
	     #Wartungszähler_Positionierachse_Zyklen(Zyklen_soll:="HMI_Wartungszähler".Wartungszähler_Positionierachse_Zyklen.Zyklen_soll,
	                                             Zyklus_Impuls:= "POS3_0_Antriebe_DB"."-1001T1_Oriental".Outputdata_FixedIO_PLC2Drv.TRIG,
	                                             Zähler_reset:="HMI_Wartungszähler".Wartungszähler_Positionierachse_Zyklen.Zähler_reset,
	                                             Zyklen_seit_Wartung=>"HMI_Wartungszähler".Wartungszähler_Positionierachse_Zyklen.Zyklen_seit_Wartung,
	                                             Zyklen_bis_Wartung=>"HMI_Wartungszähler".Wartungszähler_Positionierachse_Zyklen.Zyklen_bis_Wartung,
	                                             Gesamtzyklen=>"HMI_Wartungszähler".Wartungszähler_Positionierachse_Zyklen.Gesamtzyklen,
	                                             SM_Wartung_fällig=>"HMI_Wartungszähler".Wartungszähler_Positionierachse_Zyklen.SM_Wartung_fällig);
	    
	    IF "HMI_Wartungszähler".Wartungszähler_Positionierachse_Zyklen.Zähler_reset THEN
	        "HMI_Wartungszähler".Wartungszähler_Positionierachse_Zyklen.Zähler_reset := false;
	    END_IF;
	   
	END_REGION
	
	
	REGION Drehachse Zyklen
	    
	    
	    #Wartungszähler_Drehachse_Zyklen(Zyklen_soll := "HMI_Wartungszähler".Wartungszähler_Drehachse_Zyklen.Zyklen_soll,
	                                     Zyklus_Impuls := "POS3_0_Antriebe_DB"."-1002T2_Oriental_Drehachse".Outputdata_FixedIO_PLC2Drv.TRIG,
	                                     Zähler_reset := "HMI_Wartungszähler".Wartungszähler_Drehachse_Zyklen.Zähler_reset,
	                                     Zyklen_seit_Wartung => "HMI_Wartungszähler".Wartungszähler_Drehachse_Zyklen.Zyklen_seit_Wartung,
	                                     Zyklen_bis_Wartung => "HMI_Wartungszähler".Wartungszähler_Drehachse_Zyklen.Zyklen_bis_Wartung,
	                                     Gesamtzyklen => "HMI_Wartungszähler".Wartungszähler_Drehachse_Zyklen.Gesamtzyklen,
	                                     SM_Wartung_fällig => "HMI_Wartungszähler".Wartungszähler_Drehachse_Zyklen.SM_Wartung_fällig);
	    
	    IF "HMI_Wartungszähler".Wartungszähler_Drehachse_Zyklen.Zähler_reset THEN
	        "HMI_Wartungszähler".Wartungszähler_Drehachse_Zyklen.Zähler_reset := false;
	    END_IF;
	    
	END_REGION
	
	
	REGION Positionierachse Weg
	    IF "POS3_0_Antriebe_DB"."-1001T1_Oriental".Outputdata_FixedIO_PLC2Drv.TRIG THEN
	        #Positionierachse_Weg := ABS(("POS3_0_Antriebe_DB"."-1001T1_Oriental".Outputdata_DDO.DDO_Pos - "POS3_0_Antriebe_DB"."-1001T1_Oriental".MonitorData.FBposition) / 100);
	    END_IF;
	    
	   
	    #Wartungszähler_Positionierachse_Weg(Weg_soll := "HMI_Wartungszähler".Wartungszähler_Positionierachse_Weg.Weg_soll,
	                                         Zyklus_Impuls := "POS3_0_Antriebe_DB"."-1001T1_Oriental".Outputdata_FixedIO_PLC2Drv.TRIG,
	                                         Weg_pro_Impuls := #Positionierachse_Weg,
	                                         Zähler_reset := "HMI_Wartungszähler".Wartungszähler_Positionierachse_Weg.Zähler_reset,
	                                         Weg_seit_Wartung => "HMI_Wartungszähler".Wartungszähler_Positionierachse_Weg.Weg_seit_Wartung,
	                                         Weg_bis_Wartung => "HMI_Wartungszähler".Wartungszähler_Positionierachse_Weg.Weg_bis_Wartung,
	                                         Gesamtweg => "HMI_Wartungszähler".Wartungszähler_Positionierachse_Weg.Gesamtweg,
	                                         SM_Wartung_fällig => "HMI_Wartungszähler".Wartungszähler_Positionierachse_Weg.SM_Wartung_fällig);
	    
	    
	    
	    IF "HMI_Wartungszähler".Wartungszähler_Positionierachse_Weg.Zähler_reset THEN
	        "HMI_Wartungszähler".Wartungszähler_Positionierachse_Weg.Zähler_reset := false;
	    END_IF;
	    
	END_REGION
	
	
	REGION Drehachse Weg
	    IF "POS3_0_Antriebe_DB"."-1002T2_Oriental_Drehachse".Outputdata_FixedIO_PLC2Drv.TRIG THEN
	        #Drehachse_Weg := ABS(("POS3_0_Antriebe_DB"."-1002T2_Oriental_Drehachse".Outputdata_DDO.DDO_Pos - "POS3_0_Antriebe_DB"."-1002T2_Oriental_Drehachse".MonitorData.FBposition) / 100);
	    END_IF;
	    
	    #Wartungszähler_Drehachse_Weg(Weg_soll := "HMI_Wartungszähler".Wartungszähler_Drehachse_Weg.Weg_soll,
	                                  Zyklus_Impuls := "POS3_0_Antriebe_DB"."-1002T2_Oriental_Drehachse".Outputdata_FixedIO_PLC2Drv.TRIG,
	                                  Weg_pro_Impuls := #Drehachse_Weg,
	                                  Zähler_reset := "HMI_Wartungszähler".Wartungszähler_Drehachse_Weg.Zähler_reset,
	                                  Weg_seit_Wartung => "HMI_Wartungszähler".Wartungszähler_Drehachse_Weg.Weg_seit_Wartung,
	                                  Weg_bis_Wartung => "HMI_Wartungszähler".Wartungszähler_Drehachse_Weg.Weg_bis_Wartung,
	                                  Gesamtweg => "HMI_Wartungszähler".Wartungszähler_Drehachse_Weg.Gesamtweg,
	                                  SM_Wartung_fällig => "HMI_Wartungszähler".Wartungszähler_Drehachse_Weg.SM_Wartung_fällig);
	    
	    IF "HMI_Wartungszähler".Wartungszähler_Drehachse_Weg.Zähler_reset THEN
	        "HMI_Wartungszähler".Wartungszähler_Drehachse_Weg.Zähler_reset := false;
	    END_IF;
	    
	END_REGION
	
	
END_FUNCTION_BLOCK

FUNCTION_BLOCK "FB_Wartungszähler_Zyklen"
{ S7_Optimized_Access := 'TRUE' }
VERSION : 0.1
   VAR_INPUT 
      Zyklen_soll : DInt;
      Zyklus_Impuls : Bool;
      Zähler_reset : Bool;
   END_VAR

   VAR_OUTPUT 
      Zyklen_seit_Wartung : DInt;
      Zyklen_bis_Wartung : DInt;
      Gesamtzyklen : DInt;
      SM_Wartung_fällig : Bool;
   END_VAR

   VAR 
      R_TRIG_Zyklus_Impuls {InstructionName := 'R_TRIG'; LibVersion := '1.0'; S7_SetPoint := 'False'} : R_TRIG;
   END_VAR


BEGIN
	
	// Wartungszähler zurücksetzen
	IF #Zähler_reset THEN
	    #Zyklen_seit_Wartung := 0;
	END_IF;
	
	// Positive Flanke des Zyklusimpulses auswerten
	#R_TRIG_Zyklus_Impuls(CLK := #Zyklus_Impuls);
	
	
	IF #R_TRIG_Zyklus_Impuls.Q THEN
	    #Gesamtzyklen := #Gesamtzyklen + 1;
	    #Zyklen_seit_Wartung := #Zyklen_seit_Wartung + 1;
	END_IF;
	
	
	// Restzyklen berechnen
	IF #Zyklen_seit_Wartung < #Zyklen_soll THEN
	    #Zyklen_bis_Wartung := #Zyklen_soll - #Zyklen_seit_Wartung;
	ELSE
	    #Zyklen_bis_Wartung := 0;
	END_IF;
	
	// Wartungsmeldung setzen
	#SM_Wartung_fällig := (#Zyklen_seit_Wartung >= #Zyklen_soll);
	
END_FUNCTION_BLOCK

FUNCTION_BLOCK "FB_Wartungszähler_Weg"
{ S7_Optimized_Access := 'TRUE' }
VERSION : 0.1
   VAR_INPUT RETAIN
      Weg_soll : DInt;
      Zyklus_Impuls : Bool;
      Weg_pro_Impuls : DInt;
      Zähler_reset : Bool;
   END_VAR

   VAR_OUTPUT RETAIN
      Weg_seit_Wartung : DInt;
      Weg_bis_Wartung : DInt;
      Gesamtweg : DInt;
      SM_Wartung_fällig : Bool;
   END_VAR

   VAR 
      R_TRIG_Zyklus_Impuls {InstructionName := 'R_TRIG'; LibVersion := '1.0'; S7_SetPoint := 'False'} : R_TRIG;
   END_VAR


BEGIN
	
	// Wartungszähler zurücksetzen
	IF #Zähler_reset THEN
	    #Weg_seit_Wartung := 0;
	END_IF;
	
	// Positive Flanke des Zyklusimpulses auswerten
	#R_TRIG_Zyklus_Impuls(CLK := #Zyklus_Impuls);
	
	
	IF #R_TRIG_Zyklus_Impuls.Q THEN
	    #Gesamtweg := #Gesamtweg + #Weg_pro_Impuls;
	    #Weg_seit_Wartung := #Weg_seit_Wartung + #Weg_pro_Impuls;
	END_IF;
	
	
	// Restzyklen berechnen
	// IF #Weg_seit_Wartung < #Weg_soll THEN
	     #Weg_bis_Wartung := #Weg_soll - #Weg_seit_Wartung;
	// ELSE
	//     #Weg_bis_Wartung := 0;
	// END_IF;
	
	// Wartungsmeldung setzen
	#SM_Wartung_fällig := (#Weg_seit_Wartung >= #Weg_soll);
	
END_FUNCTION_BLOCK

FUNCTION "POS3_0_Bausteinaufrufe" : Void   // FC27, STL
{ S7_Optimized_Access := 'TRUE' }
BEGIN

NETWORK
TITLE = 

      CALL  "POS3_0_Betriebsart";

      CALL  "POS3_0_Antriebe", "POS3_0_Antriebe_DB";

      CALL  "POS3_0_Melden_Visu", "POS3_0_Melden_Visu_DB";
      CALL  "POS3_0_Teileauswertung";

      CALL  "POS3_0_Messtechnik", "POS3_0_Messtechnik_DB";




NETWORK
TITLE = 

      A     "03_Betriebsart_DB".ACK_Taste;
      =     "POS3_0_Signal".Schrittkette.ACK_EF;



      CALL  "POS3_0_SK_Ablauf", "POS3_0_SK_Ablauf_DB"
      ( OFF_SQ         := "POS3_0_Signal".Schrittkette.OFF_SQ,
        INIT_SQ        := "POS3_0_Signal".Schrittkette.INIT_SQ,
        ACK_EF         := "POS3_0_Signal".Schrittkette.ACK_EF,
        REG_EF         := ,
        ACK_S          := ,
        REG_S          := ,
        HALT_SQ        := "POS3_0_Signal".Schrittkette.HALT_SQ,
        HALT_TM        := "POS3_0_Signal".Schrittkette.HALT_TM,
        ZERO_OP        := "POS3_0_Signal".Schrittkette.ZERO_OP,
        EN_IL          := "POS3_0_Signal".Schrittkette.EN_IL,
        EN_SV          := "POS3_0_Signal".Schrittkette.EN_SV,
        EN_ACKREQ      := ,
        EN_SSKIP       := ,
        DISP_SACT      := ,
        DISP_SEF       := ,
        DISP_SALL      := ,
        S_PREV         := "POS3_0_Signal".Schrittkette.S_PREV,
        S_NEXT         := "POS3_0_Signal".Schrittkette.S_NEXT,
        SW_AUTO        := "POS3_0_Signal".Schrittkette.SW_AUTO,
        SW_TAP         := "POS3_0_Signal".Schrittkette.SW_TAP,
        SW_TOP         := 0,
        SW_MAN         := "POS3_0_Signal".Schrittkette.SW_MAN,
        S_SEL          := "POS3_0_Signal".Schrittkette.S_SEL,
        S_SELOK        := ,
        S_ON           := "POS3_0_Signal".Schrittkette.S_ON,
        S_OFF          := "POS3_0_Signal".Schrittkette.S_OFF,
        T_PREV         := ,
        T_NEXT         := ,
        T_PUSH         := "POS3_0_Signal".Schrittkette.T_PUSH,
        EN_LMODE       := ,
        S_NO           := "POS3_0_Signal".Schrittkette.S_NO,
        S_MORE         := "POS3_0_Signal".Schrittkette.S_MORE,
        S_ACTIVE       := "POS3_0_Signal".Schrittkette.S_ACTIVE,
        S_TIME         := ,
        S_TIMEOK       := ,
        S_CRITLOC      := ,
        S_CRITLOCERR   := ,
        S_STATE        := ,
        T_NO           := ,
        T_MORE         := ,
        T_CRIT         := ,
        T_CRITOLD      := ,
        T_CRITFLT      := ,
        ERROR          := ,
        FAULT          := ,
        ERR_FLT        := "POS3_0_Signal".Schrittkette.ERR_FLT,
        SQ_ISOFF       := ,
        SQ_HALTED      := "POS3_0_Signal".Schrittkette.SQ_HALTED,
        TM_HALTED      := "POS3_0_Signal".Schrittkette.TM_HALTED,
        OP_ZEROED      := "POS3_0_Signal".Schrittkette.OP_ZEROED,
        IL_ENABLED     := "POS3_0_Signal".Schrittkette.IL_ENABELD,
        SV_ENABLED     := "POS3_0_Signal".Schrittkette.SV_ENABELD,
        ACKREQ_ENABLED := ,
        SSKIP_ENABLED  := ,
        SACT_DISP      := ,
        SEF_DISP       := ,
        SALL_DISP      := ,
        AUTO_ON        := "POS3_0_Signal".Schrittkette.AUTO_ON,
        TAP_ON         := "POS3_0_Signal".Schrittkette.TAP_ON,
        TOP_ON         := ,
        MAN_ON         := "POS3_0_Signal".Schrittkette.MAN_ON,
        LMODE_ENABLED  := 
      );


END_FUNCTION

FUNCTION "POS3_0_Betriebsart" : Void   // FC40, STL
{ S7_Optimized_Access := 'TRUE' }
BEGIN

NETWORK
TITLE = Schrittkette Halt von Betriebsart
      A(;
      A     "03_Betriebsart_DB".BA_Manuell;
      A(;
      L     "HMI_SYS"."Aktueller Bildschirm";
      L     21300;  // Bildschirm Einzelschritt ist aktiv
      ==I;
      );
      );

      O     "03_Betriebsart_DB".BA_Automatik;

      O(;  // Richten aktiv oder angefordert
      A     "03_Betriebsart_DB".BA_Richten;
      A(;
      A     "POS3_0_Signal".Station.SK_Richten_gestartet;
      O     "POS3_0_Signal".Station.SK_Freigabe_Richten;
      );
      );
      NOT;
      =     "POS3_0_Signal".Station.SK_Halt_von_Betriebsart;


NETWORK
TITLE = Schrittkettenaufruf
      ON    "03_Betriebsart_DB"."NOT-HALT OK";
      ON    "03_Betriebsart_DB"."Schutztüren OK";
      O     "03_Betriebsart_DB".BA_0;
      O     "POS3_0_Signal".Station.SK_Halt_von_Betriebsart;
      AN    "POS3_0_Signal".Schrittkette.SQ_HALTED;
      A     "Zyklisch wechselnder Merker";
      O(;
      A     "03_Betriebsart_DB"."NOT-HALT OK";
      A     "03_Betriebsart_DB"."Schutztüren OK";
      AN    "03_Betriebsart_DB".BA_0;
      AN    "POS3_0_Signal".Station.SK_Halt_von_Betriebsart;
      A     "POS3_0_Signal".Schrittkette.SQ_HALTED;
      A     "Zyklisch wechselnder Merker";
      );
      =     "POS3_0_Signal".Schrittkette.HALT_SQ;

      AN    "03_Betriebsart_DB"."NOT-HALT OK";
      ON    "03_Betriebsart_DB"."Schutztüren OK";
      O     "03_Betriebsart_DB".BA_0;
      O     "POS3_0_Signal".Station.SK_Halt_von_Betriebsart;
      AN    "POS3_0_Signal".Schrittkette.TM_HALTED;
      A     "Zyklisch wechselnder Merker";
      O(;
      A     "03_Betriebsart_DB"."NOT-HALT OK";
      A     "03_Betriebsart_DB"."Schutztüren OK";
      AN    "03_Betriebsart_DB".BA_0;
      AN    "POS3_0_Signal".Station.SK_Halt_von_Betriebsart;
      A     "POS3_0_Signal".Schrittkette.TM_HALTED;
      A     "Zyklisch wechselnder Merker";
      );
      =     "POS3_0_Signal".Schrittkette.HALT_TM;

      ON    "03_Betriebsart_DB"."NOT-HALT OK";
      ON    "03_Betriebsart_DB"."Schutztüren OK";
      O     "03_Betriebsart_DB".BA_0;
      O     "POS3_0_Signal".Station.SK_Halt_von_Betriebsart;
      AN    "POS3_0_Signal".Schrittkette.OP_ZEROED;
      A     "Zyklisch wechselnder Merker";
      O(;
      A     "03_Betriebsart_DB"."NOT-HALT OK";
      A     "03_Betriebsart_DB"."Schutztüren OK";
      AN    "03_Betriebsart_DB".BA_0;
      AN    "POS3_0_Signal".Station.SK_Halt_von_Betriebsart;
      A     "POS3_0_Signal".Schrittkette.OP_ZEROED;
      A     "Zyklisch wechselnder Merker";
      );
      =     "POS3_0_Signal".Schrittkette.ZERO_OP;





NETWORK
TITLE = Tipp/Autobetriebbetrieb
      A     "HMI_BETR_ART_POS".POS3_0.Taster_Anwahl_Tipp;
      AN    "POS3_0_Signal".Schrittkette.TAP_ON;
      A     "Zyklisch wechselnder Merker";
      =     "POS3_0_Signal".Schrittkette.SW_TAP;


      AN    "HMI_BETR_ART_POS".POS3_0.Taster_Anwahl_Tipp;
      AN    "POS3_0_Signal".Schrittkette.AUTO_ON;
      A     "Zyklisch wechselnder Merker";
      =     "POS3_0_Signal".Schrittkette.SW_AUTO;

NETWORK
TITLE = Tippen
      A     "03_Betriebsart_DB".Start_Taste_FP;
      O     "HMI_BETR_ART_POS".POS3_0.Taster_Tipp_Plus;
      =     "POS3_0_Signal".Schrittkette.T_PUSH;




NETWORK
TITLE = Tippen angewählt
END_FUNCTION

FUNCTION_BLOCK "POS3_0_Antriebe"   // FB34, FBD
{ S7_Optimized_Access := 'TRUE' }
// stored: MemoryReserve 100, SetENOAutomatically false
   VAR
      "-1001T1_OM_PRM_Access_Instance" { S7_SetPoint := 'True'} : "OM_PRM_Access";
      "-1001T1_Oriental" { S7_SetPoint := 'True'} : "Oriental_AZD-KPN_Profinet";
      "-1002T2_OM_PRM_Access_Instance" { S7_SetPoint := 'True'} : "OM_PRM_Access";
      "-1002T2_Oriental_Drehachse" { S7_SetPoint := 'True'} : "Oriental_AZD-KPN_Profinet";
      Pos_Alt { S7_SetPoint := 'True'} : Real;
      Delta : Real;
   END_VAR
BEGIN

REGION Network 1 (SCL): -1001T1 Pos 3.0 Positionierachse Vorgaben Geschwindigkeit und Beschleunigung
   "POS3_0_Signal"."-1001T1 Oriental_Beschleunigung" := 50.0;
   "POS3_0_Signal"."-1001T1 Oriental_Speed" := 100.0;
END_REGION

REGION Network 2 (SCL): -1001T1 Pos 3.0 Positionierachse Achse stopp
   // Achse stopp
   IF "03_Betriebsart_DB"."Schutztüren OK" AND
       "DE_POS3_0_Endlage_Überlastzylinder" THEN
       "POS3_0_Signal"."-1001T1 Oriental_Steuerung".E_STOP := FALSE;
   ELSE
       "POS3_0_Signal"."-1001T1 Oriental_Steuerung".E_STOP := TRUE;
   END_IF;
END_REGION

REGION Network 3 (SCL): -1001T1 Pos 3.0 Positionierachse Position 0 Achse [Grundstellung]
   "POS3_0_Signal"."-1001T1 Oriental_Positionen".Operation_type[0] := 16#0001;
   "POS3_0_Signal"."-1001T1 Oriental_Positionen".Soll_Position[0] := 0.0;
   "POS3_0_Signal"."-1001T1 Oriental_Positionen".Geschwindigkeit[0] := 10.0;
   "POS3_0_Signal"."-1001T1 Oriental_Positionen".Start_Rampe[0] := "POS3_0_Signal"."-1001T1 Oriental_Beschleunigung"; // Start-Rampe %
   "POS3_0_Signal"."-1001T1 Oriental_Positionen".Stopp_Rampe[0] := "POS3_0_Signal"."-1001T1 Oriental_Beschleunigung"; // Stopp-Rampe %
   "POS3_0_Signal"."-1001T1 Oriental_Positionen".Arbeitsstrom[0] := 100;  // Arbeitsstrom in %
   "POS3_0_Signal"."-1001T1 Oriental_Positionen".Positioniertoleranz[0] := 0.02;
END_REGION

REGION Network 4 (SCL): -1001T1 Pos 3.0 Positionierachse Position 1 Achse [GS aus Verwaltung]
   "POS3_0_Signal"."-1001T1 Oriental_Positionen".Operation_type[1] := 16#0001;

   "POS3_0_Signal"."-1001T1 Oriental_Positionen".Start_Rampe[1] := "POS3_0_Signal"."-1001T1 Oriental_Beschleunigung"; // Start-Rampe %
   "POS3_0_Signal"."-1001T1 Oriental_Positionen".Stopp_Rampe[1] := "POS3_0_Signal"."-1001T1 Oriental_Beschleunigung"; // Stopp-Rampe %
   "POS3_0_Signal"."-1001T1 Oriental_Positionen".Arbeitsstrom[1] := 100;   // Arbeitsstrom in %
   "POS3_0_Signal"."-1001T1 Oriental_Positionen".Positioniertoleranz[1] := 0.02;
END_REGION

REGION Network 5 (SCL): -1001T1 Pos 3.0 Positionierachse Position 2 Achse [AS aus Verwaltung]
   "POS3_0_Signal"."-1001T1 Oriental_Positionen".Operation_type[2] := 16#0001;

   "POS3_0_Signal"."-1001T1 Oriental_Positionen".Start_Rampe[2] := "POS3_0_Signal"."-1001T1 Oriental_Beschleunigung"; // Start-Rampe %
   "POS3_0_Signal"."-1001T1 Oriental_Positionen".Stopp_Rampe[2] := "POS3_0_Signal"."-1001T1 Oriental_Beschleunigung"; // Stopp-Rampe %
   "POS3_0_Signal"."-1001T1 Oriental_Positionen".Arbeitsstrom[2] := 100;  // Arbeitsstrom in %
   "POS3_0_Signal"."-1001T1 Oriental_Positionen".Positioniertoleranz[2] := 0.02;
END_REGION

REGION Network 6 (SCL): -1001T1 Pos 3.0 Positionierachse Position 3 Achse
   "POS3_0_Signal"."-1001T1 Oriental_Positionen".Operation_type[3] := 16#0001;

   "POS3_0_Signal"."-1001T1 Oriental_Positionen".Start_Rampe[3] := "POS3_0_Signal"."-1001T1 Oriental_Beschleunigung" ; // Start-Rampe %
   "POS3_0_Signal"."-1001T1 Oriental_Positionen".Stopp_Rampe[3] := "POS3_0_Signal"."-1001T1 Oriental_Beschleunigung" ; // Stopp-Rampe %
   "POS3_0_Signal"."-1001T1 Oriental_Positionen".Arbeitsstrom[3] := 100; // Arbeitsstrom in %
   "POS3_0_Signal"."-1001T1 Oriental_Positionen".Positioniertoleranz[3] := 0.02;
END_REGION

REGION Network 7 (SCL): -1001T1 Pos 3.0 Positionierachse Position 4 Achse
   "POS3_0_Signal"."-1001T1 Oriental_Positionen".Operation_type[4] := 16#0001;

   "POS3_0_Signal"."-1001T1 Oriental_Positionen".Start_Rampe[4] := "POS3_0_Signal"."-1001T1 Oriental_Beschleunigung" ; // Start-Rampe %
   "POS3_0_Signal"."-1001T1 Oriental_Positionen".Stopp_Rampe[4] := "POS3_0_Signal"."-1001T1 Oriental_Beschleunigung" ; // Stopp-Rampe %
   "POS3_0_Signal"."-1001T1 Oriental_Positionen".Arbeitsstrom[4] := 100;  // Arbeitsstrom in %
   "POS3_0_Signal"."-1001T1 Oriental_Positionen".Positioniertoleranz[4] := 0.03;
END_REGION

REGION Network 8 (SCL): -1001T1 Pos 3.0 Positionierachse Position 5 Achse

   "POS3_0_Signal"."-1001T1 Oriental_Positionen".Operation_type[5] := 16#0001;

   "POS3_0_Signal"."-1001T1 Oriental_Positionen".Start_Rampe[5] := "POS3_0_Signal"."-1001T1 Oriental_Beschleunigung"; // Start-Rampe %
   "POS3_0_Signal"."-1001T1 Oriental_Positionen".Stopp_Rampe[5] := "POS3_0_Signal"."-1001T1 Oriental_Beschleunigung"; // Stopp-Rampe %
   "POS3_0_Signal"."-1001T1 Oriental_Positionen".Arbeitsstrom[5] := 100;  // Arbeitsstrom in %
   "POS3_0_Signal"."-1001T1 Oriental_Positionen".Positioniertoleranz[5] := 0.03;
END_REGION

REGION Network 9 (SCL): -1001T1 Pos 3.0 Positionierachse Grenzwerte
   "POS3_0_Signal"."-1001T1 Oriental_Positionen".A_Softw_ES_max_mm := 210.0;
   "POS3_0_Signal"."-1001T1 Oriental_Positionen".A_Softw_ES_min_mm := -0.5;
END_REGION

NETWORK
TITLE = -1001T1 Pos 3.0 Positionierachse E_ETO-CLR Quittieren nach "Sicherer Halt"
      A     "03_Betriebsart_DB"."NOT-HALT OK";
      A     "03_Betriebsart_DB"."Schutztüren OK";
      AN    "POS3_0_Signal"."-1001T1 Oriental_Steuerung"."A_DCMD-RDY";
      A     "FL_Clock_1Hz";
      =     "POS3_0_Signal"."-1001T1 Oriental_Steuerung"."E_ETO-CLR";


NETWORK
TITLE = -1001T1 Pos 3.0 Positionierachse Oriental Achse Parameter schreiben und lesen (wird nicht benötigt)
      CALL  #"-1001T1_OM_PRM_Access_Instance"
      ( Inputdata_RW_Drv2PLC  := "AZ_1001T1_Pos3_0__Prm_Status",
        ReadParameterID       := "POS3_0_Parameter_Data".RD_ParameterID,
        WriteParameterID      := "POS3_0_Parameter_Data".WR_ParameterID,
        WriteData             := "POS3_0_Parameter_Data".WR_ParameterData,
        "WR-REQ"              := ,
        Outputdata_RW_PLC2Drv := "AZ_1001T1_Pos3_0__Prm_Set",
        ReadParameterID_R     := ,
        WriteParameterID_R    := ,
        ReadData              := "POS3_0_Parameter_Data".RD_ParameterData,
        "WR-SET-ERR"          := ,
        "WR-IF-ERR"           := ,
        "WR-NV-ERR"           := ,
        "WR-EXE-ERR"          := ,
        "WR-ERR"              := ,
        "RD-ERR"              := ,
        "WR-END"              := ,
        "SYS-BSY"             := 
      );



REGION Network 12 (SCL): -1001T1 Pos 3.0 Positionierachse Oriental DDO_Type für E_Trig_Manuell
   // E_DDO_Type 16#0001 = absolut positionieren 16#0002 = relativ positionieren
   "POS3_0_Signal"."-1001T1 Oriental_Steuerung".E_DDO_Type := 16#0001;
END_REGION

NETWORK
TITLE = -1001T1 Pos 3.0 Positionierachse Oriental Achse Ansteuerung
      CALL  #"-1001T1_Oriental"
      ( Inputdata_FixedIO_Drv2PLC           := "AZ_1001T1_Pos3_0__Fixed_Out",
        MonitorData                         := "AZ_1001T1_Pos3_0__St_Monitor",
        E_DDO_Type                          := "POS3_0_Signal"."-1001T1 Oriental_Steuerung".E_DDO_Type,
        E_DDO_Pos                           := "POS3_0_Signal"."-1001T1 Oriental_Steuerung".E_DDO_Pos,
        E_DDO_Vel                           := "POS3_0_Signal"."-1001T1 Oriental_Steuerung".E_DDO_Vel,
        E_DDO_Acc                           := "POS3_0_Signal"."-1001T1 Oriental_Steuerung".E_DDO_Acc,
        E_DDO_Dec                           := "POS3_0_Signal"."-1001T1 Oriental_Steuerung".E_DDO_Dec,
        E_DDO_Crnt                          := "POS3_0_Signal"."-1001T1 Oriental_Steuerung".E_DDO_Crnt,
        E_DDO_Trans                         := "POS3_0_Signal"."-1001T1 Oriental_Steuerung".E_DDO_Trans,
        E_Schrittweite_Pos                  := "POS3_0_Signal"."-1001T1 Oriental_Steuerung".E_Schrittweite_pos,
        E_Schrittweite_Neg                  := "POS3_0_Signal"."-1001T1 Oriental_Steuerung".E_Schrittweite_neg,
        E_Schrittweite                      := "POS3_0_Signal"."-1001T1 Oriental_Steuerung".E_Schrittweite,
        E_R_Softw_ES_min_steps              := "POS3_0_Signal"."-1001T1 Oriental_Positionen".A_Softw_ES_min_mm,
        E_R_Softw_ES_max_steps              := "POS3_0_Signal"."-1001T1 Oriental_Positionen".A_Softw_ES_max_mm,
        E_Drehachse                         := FALSE,
        E_Getriebefaktor                    := 100.0,
        E_Maximalgeschwindigkeit_Hz         := 25000.0,
        "E_Maximal_Start_Stopp_Rampe_kHz/s" := 250000.0,
        E_SIMULATION_AKTIV                  := "03_Betriebsart_DB".Simulation_aktiv,
        E_RemoteIO                          := "AZ_1001T1_Pos3_0__Remote_Out",
        Outputdata_DDO                      := "AZ_1001T1_Pos3_0__DDO",
        Outputdata_FixedIO_PLC2Drv          := "AZ_1001T1_Pos3_0__Fixed_In",
        A_TRIG_R                            := "POS3_0_Signal"."-1001T1 Oriental_Steuerung".A_TRIG_R,
        "A_TRIG-MODE_R"                     := "POS3_0_Signal"."-1001T1 Oriental_Steuerung"."A_TRIG-MODE_R",
        "A_SET-ERR"                         := "POS3_0_Signal"."-1001T1 Oriental_Steuerung"."A_SET-ERR",
        "A_EXE-ERR"                         := "POS3_0_Signal"."-1001T1 Oriental_Steuerung"."A_EXE-ERR",
        "A_DCMD-FULL"                       := "POS3_0_Signal"."-1001T1 Oriental_Steuerung"."A_DCMD-FULL",
        A_STOP_R                            := "POS3_0_Signal"."-1001T1 Oriental_Steuerung".A_STOP_R,
        "A_ETO-MON"                         := "POS3_0_Signal"."-1001T1 Oriental_Steuerung"."A_ETO-MON",
        A_TLC                               := "POS3_0_Signal"."-1001T1 Oriental_Steuerung".A_TLC,
        "A_SEQ-BSY"                         := "POS3_0_Signal"."-1001T1 Oriental_Steuerung"."A_SEQ-BSY",
        A_MOVE                              := "POS3_0_Signal"."-1001T1 Oriental_Steuerung".A_MOVE,
        "A_IN-POS"                          := "POS3_0_Signal"."-1001T1 Oriental_Steuerung"."A_IN-POS",
        A_START_R                           := "POS3_0_Signal"."-1001T1 Oriental_Steuerung".A_START_R,
        "A_HOME-END"                        := "POS3_0_Signal"."-1001T1 Oriental_Steuerung"."A_HOME-END",
        A_READY                             := "POS3_0_Signal"."-1001T1 Oriental_Steuerung".A_READY,
        "A_DCMD-RDY"                        := "POS3_0_Signal"."-1001T1 Oriental_Steuerung"."A_DCMD-RDY",
        "A_ALM-A"                           := "POS3_0_Signal"."-1001T1 Oriental_Steuerung"."A_ALM-A",
        A_PresentAlarm                      := "POS3_0_Signal"."-1001T1 Oriental_Steuerung".A_PresentAlarm,
        A_FBposition                        := "POS3_0_Signal"."-1001T1 Oriental_Steuerung".A_FBposition,
        A_FBspeed                           := "POS3_0_Signal"."-1001T1 Oriental_Steuerung".A_FBspeed,
        A_CmdPosition                       := "POS3_0_Signal"."-1001T1 Oriental_Steuerung".A_CmdPosition,
        A_TorqueMonitor                     := "POS3_0_Signal"."-1001T1 Oriental_Steuerung".A_TorqueMonitor,
        A_CST_OpeCurrent                    := "POS3_0_Signal"."-1001T1 Oriental_Steuerung".A_CST_OpeCurrent,
        A_Information                       := "POS3_0_Signal"."-1001T1 Oriental_Steuerung".A_Information,
        A_StatusWord                        := "POS3_0_Signal"."-1001T1 Oriental_Steuerung".A_StatusWord,
        A_RemoteIO                          := "AZ_1001T1_Pos3_0__Remote_IN",
        E_A_UDT_Positionen                  := "POS3_0_Signal"."-1001T1 Oriental_Positionen",
        E_Not_Aus_OK                        := "03_Betriebsart_DB"."NOT-HALT OK",
        E_Tueren_OK                         := "03_Betriebsart_DB"."Schutztüren OK",
        "E_TRIG-MODE"                       := "POS3_0_Signal"."-1001T1 Oriental_Steuerung"."E_TRIG-MODE",
        "E_ETO-CLR"                         := "POS3_0_Signal"."-1001T1 Oriental_Steuerung"."E_ETO-CLR",
        "E_FW-JOG"                          := "POS3_0_Signal"."-1001T1 Oriental_Steuerung"."E_FW-JOG",
        "E_RV-JOG"                          := "POS3_0_Signal"."-1001T1 Oriental_Steuerung"."E_RV-JOG",
        E_START                             := "POS3_0_Signal"."-1001T1 Oriental_Steuerung".E_START,
        E_ZHOME                             := "POS3_0_Signal"."-1001T1 Oriental_Steuerung".E_ZHOME,
        E_STOP                              := "POS3_0_Signal"."-1001T1 Oriental_Steuerung".E_STOP,
        E_FREE                              := "POS3_0_Signal"."-1001T1 Oriental_Steuerung".E_FREE,
        "E_ALM-RST"                         := "03_Betriebsart_DB".ACK_Taste,
        E_TRIG_MANUELL                      := "POS3_0_Signal"."-1001T1 Oriental_Steuerung".E_Trig_Manuell,
        E_Home                              := "POS3_0_Signal"."-1001T1 Oriental_E_P-Preset"
      );

REGION Network 14 (SCL): -1001T1 Pos 3.0 "P-Preset" Reset
   IF "POS3_0_Signal"."-1001T1 Oriental_E_P-Preset" THEN
       "POS3_0_Signal"."-1001T1 Oriental_E_P-Preset" := False;
   END_IF;
END_REGION

REGION Network 16 (SCL): -1002T1 Pos 3.0 Drehachse Vorgaben Geschwindigkeit und Beschleunigung
   "POS3_0_Signal"."-1002T1_Oriental_Beschleunigung" := 40.0;
   "POS3_0_Signal"."-1002T1_Oriental_Speed" := 100.0;
END_REGION

REGION Network 17 (SCL): -1002T1 Pos 3.0 Drehachse Achse stopp
   // Achse stopp
   IF "03_Betriebsart_DB"."Schutztüren OK" THEN
       "POS3_0_Signal"."-1002T1 Oriental_Steuerung".E_STOP := FALSE;
   ELSE
       "POS3_0_Signal"."-1002T1 Oriental_Steuerung".E_STOP := TRUE;
   END_IF;
END_REGION

REGION Network 18 (SCL): -1002T1 Pos 3.0 Drehachse Position 0 [Grundstellung]
   "POS3_0_Signal"."-1002T1 Oriental_Positionen".Operation_type[0] := 16#0001;
   "POS3_0_Signal"."-1002T1 Oriental_Positionen".Soll_Position[0] := 0.0;
   "POS3_0_Signal"."-1002T1 Oriental_Positionen".Geschwindigkeit[0] := 10.0;
   "POS3_0_Signal"."-1002T1 Oriental_Positionen".Start_Rampe[0] := "POS3_0_Signal"."-1002T1_Oriental_Beschleunigung"; // Start-Rampe %
   "POS3_0_Signal"."-1002T1 Oriental_Positionen".Stopp_Rampe[0] := "POS3_0_Signal"."-1002T1_Oriental_Beschleunigung"; // Stopp-Rampe %
   "POS3_0_Signal"."-1002T1 Oriental_Positionen".Arbeitsstrom[0] := 100;  // Arbeitsstrom in %
   "POS3_0_Signal"."-1002T1 Oriental_Positionen".Positioniertoleranz[0] := 0.001;
END_REGION

REGION Network 19 (SCL): -1002T1 Pos 3.0 Drehachse Position 1 [0.0 ° Absolut positionieren]
   "POS3_0_Signal"."-1002T1 Oriental_Positionen".Operation_type[1] := 16#0001;
   "POS3_0_Signal"."-1002T1 Oriental_Positionen".Soll_Position[1] := 0.0;
   "POS3_0_Signal"."-1002T1 Oriental_Positionen".Geschwindigkeit[1] := 10.0;
   "POS3_0_Signal"."-1002T1 Oriental_Positionen".Start_Rampe[1] := "POS3_0_Signal"."-1002T1_Oriental_Beschleunigung"; // Start-Rampe %
   "POS3_0_Signal"."-1002T1 Oriental_Positionen".Stopp_Rampe[1] := "POS3_0_Signal"."-1002T1_Oriental_Beschleunigung"; // Stopp-Rampe %
   "POS3_0_Signal"."-1002T1 Oriental_Positionen".Arbeitsstrom[1] := 100;   // Arbeitsstrom in %
   "POS3_0_Signal"."-1002T1 Oriental_Positionen".Positioniertoleranz[1] := 0.001;
END_REGION

REGION Network 20 (SCL): -1002T1 Pos 3.0 Drehachse Position 2 [AS1 aus Verwaltung]
   "POS3_0_Signal"."-1002T1 Oriental_Positionen".Operation_type[2] := 16#0002;

   "POS3_0_Signal"."-1002T1 Oriental_Positionen".Start_Rampe[2] := "POS3_0_Signal"."-1002T1_Oriental_Beschleunigung"; // Start-Rampe %
   "POS3_0_Signal"."-1002T1 Oriental_Positionen".Stopp_Rampe[2] := "POS3_0_Signal"."-1002T1_Oriental_Beschleunigung"; // Stopp-Rampe %
   "POS3_0_Signal"."-1002T1 Oriental_Positionen".Arbeitsstrom[2] := REAL_TO_DINT ("Verwaltung_Teiledaten"."Drehantrieb Motorstrombegrenzung");  // Arbeitsstrom in %
   "POS3_0_Signal"."-1002T1 Oriental_Positionen".Positioniertoleranz[2] := 0.001;
END_REGION

REGION Network 21 (SCL): -1002T1 Pos 3.0 Drehachse Position 3 [GS aus Verwaltung]
   "POS3_0_Signal"."-1002T1 Oriental_Positionen".Operation_type[3] := 16#0002;

   "POS3_0_Signal"."-1002T1 Oriental_Positionen".Start_Rampe[3] := "POS3_0_Signal"."-1002T1_Oriental_Beschleunigung"; // Start-Rampe %
   "POS3_0_Signal"."-1002T1 Oriental_Positionen".Stopp_Rampe[3] := "POS3_0_Signal"."-1002T1_Oriental_Beschleunigung"; // Stopp-Rampe %
   "POS3_0_Signal"."-1002T1 Oriental_Positionen".Arbeitsstrom[3] := REAL_TO_DINT ("Verwaltung_Teiledaten"."Drehantrieb Motorstrombegrenzung");  // Arbeitsstrom in %
   "POS3_0_Signal"."-1002T1 Oriental_Positionen".Positioniertoleranz[3] := 0.001;
END_REGION

REGION Network 22 (SCL): -1002T1 Pos 3.0 Drehachse Position 4
   "POS3_0_Signal"."-1002T1 Oriental_Positionen".Operation_type[4] := 16#0001;

   "POS3_0_Signal"."-1002T1 Oriental_Positionen".Start_Rampe[4] := "POS3_0_Signal"."-1002T1_Oriental_Beschleunigung"; // Start-Rampe %
   "POS3_0_Signal"."-1002T1 Oriental_Positionen".Stopp_Rampe[4] := "POS3_0_Signal"."-1002T1_Oriental_Beschleunigung"; // Stopp-Rampe %
   "POS3_0_Signal"."-1002T1 Oriental_Positionen".Arbeitsstrom[4] := 100;  // Arbeitsstrom in %
   "POS3_0_Signal"."-1002T1 Oriental_Positionen".Positioniertoleranz[4] := 0.01;
END_REGION

REGION Network 23 (SCL): -1002T1 Pos 3.0 Drehachse Position 5
   "POS3_0_Signal"."-1002T1 Oriental_Positionen".Operation_type[5] := 16#0001;

   "POS3_0_Signal"."-1002T1 Oriental_Positionen".Start_Rampe[5] := "POS3_0_Signal"."-1002T1_Oriental_Beschleunigung"; // Start-Rampe %
   "POS3_0_Signal"."-1002T1 Oriental_Positionen".Stopp_Rampe[5] := "POS3_0_Signal"."-1002T1_Oriental_Beschleunigung"; // Stopp-Rampe %
   "POS3_0_Signal"."-1002T1 Oriental_Positionen".Arbeitsstrom[5] := 100;  // Arbeitsstrom in %
   "POS3_0_Signal"."-1002T1 Oriental_Positionen".Positioniertoleranz[5] := 0.01;
END_REGION

REGION Network 24 (SCL): -1002T1 Pos 3.0 Drehachse Grenzwerte
   "POS3_0_Signal"."-1002T1 Oriental_Positionen".A_Softw_ES_max_mm := 10000.5;
   "POS3_0_Signal"."-1002T1 Oriental_Positionen".A_Softw_ES_min_mm := -10000.5;
END_REGION

NETWORK
TITLE = -1002T1 Pos 3.0 Drehachse E_ETO-CLR Quittieren nach "Sicherer Halt"
      A     "03_Betriebsart_DB"."NOT-HALT OK";
      A     "03_Betriebsart_DB"."Schutztüren OK";
      AN    "POS3_0_Signal"."-1002T1 Oriental_Steuerung"."A_DCMD-RDY";
      A     "FL_Clock_1Hz";
      =     "POS3_0_Signal"."-1002T1 Oriental_Steuerung"."E_ETO-CLR";


NETWORK
TITLE = -1002T1 Pos 3.0 Drehachse Oriental Achse Parameter schreiben und lesen (wird nicht benötigt)
      CALL  #"-1002T2_OM_PRM_Access_Instance"
      ( Inputdata_RW_Drv2PLC  := "AZ_1002T1_Pos3_0_Drehachse__Prm_Status",
        ReadParameterID       := "POS3_0_Parameter_Data_Drehachse".RD_ParameterID,
        WriteParameterID      := "POS3_0_Parameter_Data_Drehachse".WR_ParameterID,
        WriteData             := "POS3_0_Parameter_Data_Drehachse".WR_ParameterData,
        "WR-REQ"              := ,
        Outputdata_RW_PLC2Drv := "AZ_1002T1_Pos3_0_Drehachse__Prm_Set",
        ReadParameterID_R     := ,
        WriteParameterID_R    := ,
        ReadData              := "POS3_0_Parameter_Data_Drehachse".RD_ParameterData,
        "WR-SET-ERR"          := ,
        "WR-IF-ERR"           := ,
        "WR-NV-ERR"           := ,
        "WR-EXE-ERR"          := ,
        "WR-ERR"              := ,
        "RD-ERR"              := ,
        "WR-END"              := ,
        "SYS-BSY"             := 
      );



REGION Network 27 (SCL): -1002T1 Pos 3.0 Drehachse DDO_Type für E_Trig_Manuell
   // E_DDO_Type 16#0001 = absolut positionieren 16#0002 = relativ positionieren
   "POS3_0_Signal"."-1002T1 Oriental_Steuerung".E_DDO_Type := 16#0002;
END_REGION

NETWORK
TITLE = -1002T1 Pos 3.0 Drehachse Oriental Achse Ansteuerung
      CALL  #"-1002T2_Oriental_Drehachse"
      ( Inputdata_FixedIO_Drv2PLC           := "AZ_1002T1_Pos3_0_Drehachse__Fixed_Out",
        MonitorData                         := "AZ_1002T1_Pos3_0_Drehachse__St_Monitor",
        E_DDO_Type                          := "POS3_0_Signal"."-1002T1 Oriental_Steuerung".E_DDO_Type,
        E_DDO_Pos                           := "POS3_0_Signal"."-1002T1 Oriental_Steuerung".E_DDO_Pos,
        E_DDO_Vel                           := "POS3_0_Signal"."-1002T1 Oriental_Steuerung".E_DDO_Vel,
        E_DDO_Acc                           := "POS3_0_Signal"."-1002T1 Oriental_Steuerung".E_DDO_Acc,
        E_DDO_Dec                           := "POS3_0_Signal"."-1002T1 Oriental_Steuerung".E_DDO_Dec,
        E_DDO_Crnt                          := "POS3_0_Signal"."-1002T1 Oriental_Steuerung".E_DDO_Crnt,
        E_DDO_Trans                         := "POS3_0_Signal"."-1002T1 Oriental_Steuerung".E_DDO_Trans,
        E_Schrittweite_Pos                  := "POS3_0_Signal"."-1002T1 Oriental_Steuerung".E_Schrittweite_pos,
        E_Schrittweite_Neg                  := "POS3_0_Signal"."-1002T1 Oriental_Steuerung".E_Schrittweite_neg,
        E_Schrittweite                      := "POS3_0_Signal"."-1002T1 Oriental_Steuerung".E_Schrittweite,
        E_R_Softw_ES_min_steps              := "POS3_0_Signal"."-1002T1 Oriental_Positionen".A_Softw_ES_min_mm,
        E_R_Softw_ES_max_steps              := "POS3_0_Signal"."-1002T1 Oriental_Positionen".A_Softw_ES_max_mm,
        E_Drehachse                         := TRUE,
        E_Getriebefaktor                    := 18.0,
        E_Maximalgeschwindigkeit_Hz         := 30000.0,
        "E_Maximal_Start_Stopp_Rampe_kHz/s" := 990000.0,
        E_SIMULATION_AKTIV                  := "03_Betriebsart_DB".Simulation_aktiv,
        E_RemoteIO                          := "AZ_1002T1_Pos3_0_Drehachse__Remote_Out",
        Outputdata_DDO                      := "AZ_1002T1_Pos3_0_Drehachse__DDO",
        Outputdata_FixedIO_PLC2Drv          := "AZ_1002T1_Pos3_0_Drehachse__Fixed_In",
        A_TRIG_R                            := "POS3_0_Signal"."-1002T1 Oriental_Steuerung".A_TRIG_R,
        "A_TRIG-MODE_R"                     := "POS3_0_Signal"."-1002T1 Oriental_Steuerung"."A_TRIG-MODE_R",
        "A_SET-ERR"                         := "POS3_0_Signal"."-1002T1 Oriental_Steuerung"."A_SET-ERR",
        "A_EXE-ERR"                         := "POS3_0_Signal"."-1002T1 Oriental_Steuerung"."A_EXE-ERR",
        "A_DCMD-FULL"                       := "POS3_0_Signal"."-1002T1 Oriental_Steuerung"."A_DCMD-FULL",
        A_STOP_R                            := "POS3_0_Signal"."-1002T1 Oriental_Steuerung".A_STOP_R,
        "A_ETO-MON"                         := "POS3_0_Signal"."-1002T1 Oriental_Steuerung"."A_ETO-MON",
        A_TLC                               := "POS3_0_Signal"."-1002T1 Oriental_Steuerung".A_TLC,
        "A_SEQ-BSY"                         := "POS3_0_Signal"."-1002T1 Oriental_Steuerung"."A_SEQ-BSY",
        A_MOVE                              := "POS3_0_Signal"."-1002T1 Oriental_Steuerung".A_MOVE,
        "A_IN-POS"                          := "POS3_0_Signal"."-1002T1 Oriental_Steuerung"."A_IN-POS",
        A_START_R                           := "POS3_0_Signal"."-1002T1 Oriental_Steuerung".A_START_R,
        "A_HOME-END"                        := "POS3_0_Signal"."-1002T1 Oriental_Steuerung"."A_HOME-END",
        A_READY                             := "POS3_0_Signal"."-1002T1 Oriental_Steuerung".A_READY,
        "A_DCMD-RDY"                        := "POS3_0_Signal"."-1002T1 Oriental_Steuerung"."A_DCMD-RDY",
        "A_ALM-A"                           := "POS3_0_Signal"."-1002T1 Oriental_Steuerung"."A_ALM-A",
        A_PresentAlarm                      := "POS3_0_Signal"."-1002T1 Oriental_Steuerung".A_PresentAlarm,
        A_FBposition                        := "POS3_0_Signal"."-1002T1 Oriental_Steuerung".A_FBposition,
        A_FBspeed                           := "POS3_0_Signal"."-1002T1 Oriental_Steuerung".A_FBspeed,
        A_CmdPosition                       := "POS3_0_Signal"."-1002T1 Oriental_Steuerung".A_CmdPosition,
        A_TorqueMonitor                     := "POS3_0_Signal"."-1002T1 Oriental_Steuerung".A_TorqueMonitor,
        A_CST_OpeCurrent                    := "POS3_0_Signal"."-1002T1 Oriental_Steuerung".A_CST_OpeCurrent,
        A_Information                       := "POS3_0_Signal"."-1002T1 Oriental_Steuerung".A_Information,
        A_StatusWord                        := "POS3_0_Signal"."-1002T1 Oriental_Steuerung".A_StatusWord,
        A_RemoteIO                          := "AZ_1002T1_Pos3_0_Drehachse__Remote_IN",
        E_A_UDT_Positionen                  := "POS3_0_Signal"."-1002T1 Oriental_Positionen",
        E_Not_Aus_OK                        := "03_Betriebsart_DB"."NOT-HALT OK",
        E_Tueren_OK                         := "03_Betriebsart_DB"."Schutztüren OK",
        "E_TRIG-MODE"                       := "POS3_0_Signal"."-1002T1 Oriental_Steuerung"."E_TRIG-MODE",
        "E_ETO-CLR"                         := "POS3_0_Signal"."-1002T1 Oriental_Steuerung"."E_ETO-CLR",
        "E_FW-JOG"                          := "POS3_0_Signal"."-1002T1 Oriental_Steuerung"."E_FW-JOG",
        "E_RV-JOG"                          := "POS3_0_Signal"."-1002T1 Oriental_Steuerung"."E_RV-JOG",
        E_START                             := "POS3_0_Signal"."-1002T1 Oriental_Steuerung".E_START,
        E_ZHOME                             := "POS3_0_Signal"."-1002T1 Oriental_Steuerung".E_ZHOME,
        E_STOP                              := "POS3_0_Signal"."-1002T1 Oriental_Steuerung".E_STOP,
        E_FREE                              := "POS3_0_Signal"."-1002T1 Oriental_Steuerung".E_FREE,
        "E_ALM-RST"                         := "03_Betriebsart_DB".ACK_Taste,
        E_TRIG_MANUELL                      := "POS3_0_Signal"."-1002T1 Oriental_Steuerung".E_Trig_Manuell,
        E_Home                              := "POS3_0_Signal"."-1002T1 Oriental_E_P-Preset"
      );

REGION Network 29 (SCL): -1002T1 Pos 3.0 Drehachse "P-Preset" Reset
   IF "POS3_0_Signal"."-1002T1 Oriental_E_P-Preset" THEN
       "POS3_0_Signal"."-1002T1 Oriental_E_P-Preset" := False;
       "POS3_0_Signal"."-1002T1 Oriental_Umdrehungszähler" := 0.0;
   END_IF;
END_REGION

REGION Network 30 (SCL): -1002T1 Pos 3.0 Drehachse Berechnung der Umdrehungen ab dem Nullpunkt
   // Positionsdifferenz berechnen
   #Delta := "POS3_0_Signal"."-1002T1 Oriental_Steuerung".A_FBposition - #Pos_Alt;

   //Überlauf erkennen 
   IF #Delta < -180.0 THEN
       // Vorwärts über 360° gelaufen (z.B. 359 -> 1)
       "POS3_0_Signal"."-1002T1 Oriental_Umdrehungszähler" :=
       "POS3_0_Signal"."-1002T1 Oriental_Umdrehungszähler" + 1.0;

   ELSIF #Delta > 180.0 THEN
       // Rückwärts über 0° gelaufen (z.B. 1 -> 359)    
       "POS3_0_Signal"."-1002T1 Oriental_Umdrehungszähler" :=
       "POS3_0_Signal"."-1002T1 Oriental_Umdrehungszähler" - 1.0;
   END_IF;

   // Aktuellen Wert für nächsten Zyklus speichern
   #Pos_Alt := "POS3_0_Signal"."-1002T1 Oriental_Steuerung".A_FBposition;


   "POS3_0_Signal"."-1002T1 Oriental_Absolute_Position" :=    "POS3_0_Signal"."-1002T1 Oriental_Umdrehungszähler" * 360.0 +
   "POS3_0_Signal"."-1002T1 Oriental_Steuerung".A_FBposition;
END_REGION

REGION Network 31 (SCL): -1002T1 Pos 3.0 Drehachse Kraft überschritten
   IF "POS3_0_Signal"."-1002T1 Oriental_Steuerung".A_TorqueMonitor >=
      "POS3_0_Signal"."-1002T1 Oriental_Steuerung".A_CST_OpeCurrent   THEN
       "POS3_0_Signal".Drehachse_Kraft_überschritten := true;
   ELSE
       "POS3_0_Signal".Drehachse_Kraft_überschritten := false;
   END_IF;
END_REGION
END_FUNCTION_BLOCK

FUNCTION_BLOCK "OM_PRM_Access"   // FB82, LAD
{ S7_Optimized_Access := 'TRUE' }
// stored: MemoryReserve 100, SetENOAutomatically false
   VAR_INPUT
      Inputdata_RW_Drv2PLC : "AZ_PrmRW_Drv2PLC";
      ReadParameterID : Word;
      WriteParameterID : Word;
      WriteData : DWord;
      "WR-REQ" : Bool;
   END_VAR
   VAR_OUTPUT
      Outputdata_RW_PLC2Drv : "AZ_PrmRW_PLC2Drv";
      ReadParameterID_R : Word;
      WriteParameterID_R : Word;
      ReadData : DWord;
      "WR-SET-ERR" : Bool;
      "WR-IF-ERR" : Bool;
      "WR-NV-ERR" : Bool;
      "WR-EXE-ERR" : Bool;
      "WR-ERR" : Bool;
      "RD-ERR" : Bool;
      "WR-END" : Bool;
      "SYS-BSY" : Bool;
   END_VAR
BEGIN

REGION Network 1
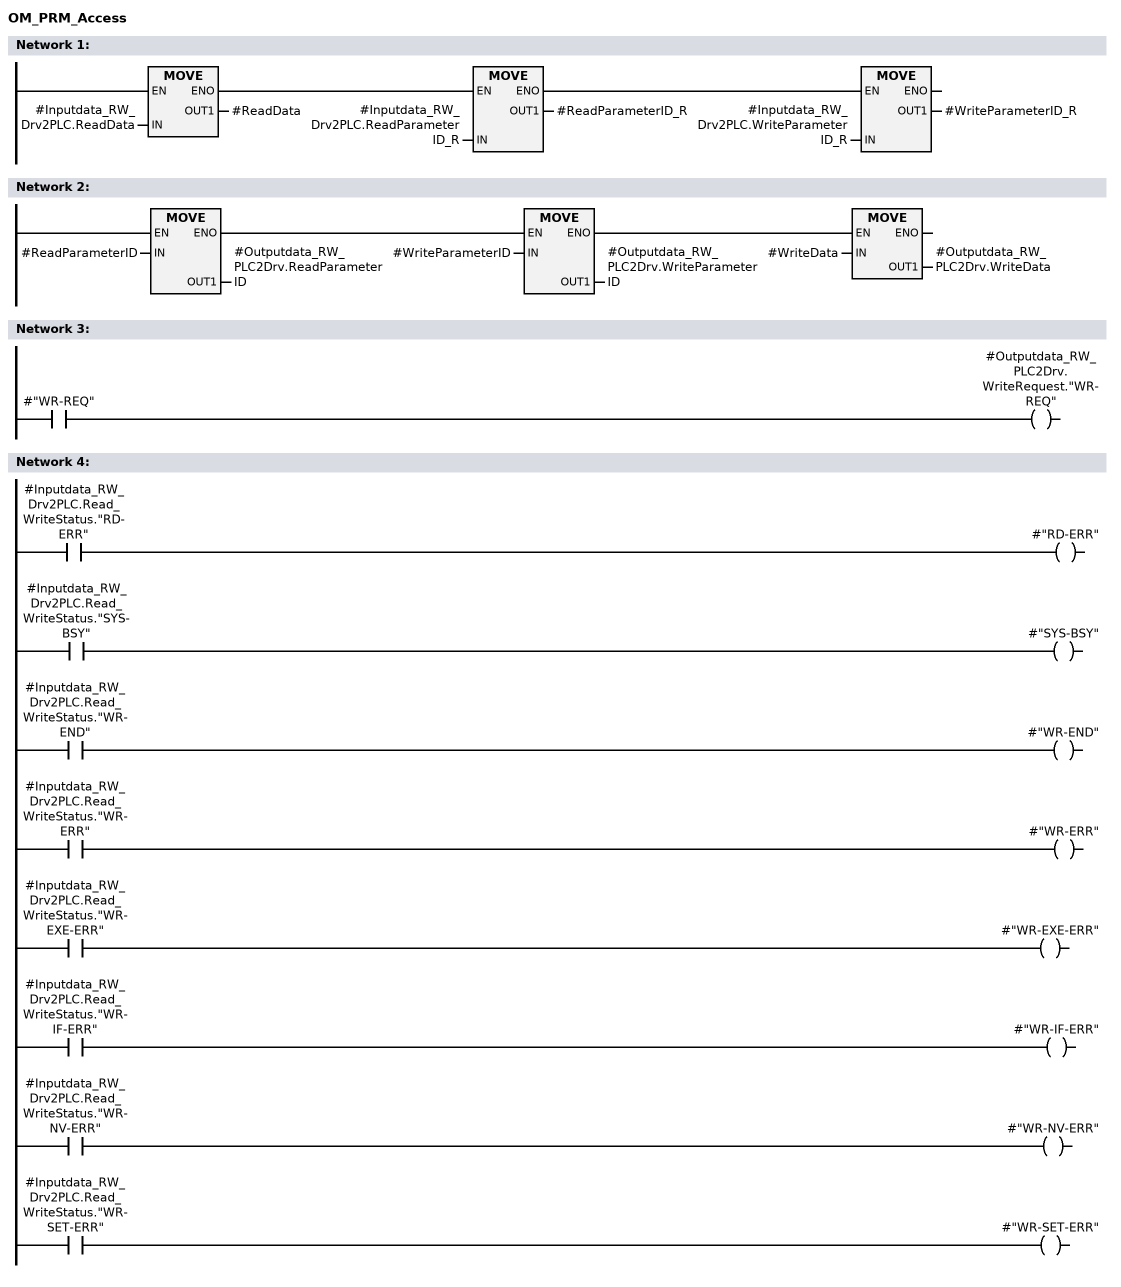
   RUNG wire#powerrail
      Move(in := #Inputdata_RW_Drv2PLC.ReadData, out1 => #ReadData)
      Move(in := #Inputdata_RW_Drv2PLC.ReadParameterID_R, out1 => #ReadParameterID_R)
      Move(in := #Inputdata_RW_Drv2PLC.WriteParameterID_R, out1 => #WriteParameterID_R)
   END_RUNG
   // the same network as SCL:
   #ReadData := #Inputdata_RW_Drv2PLC.ReadData;
   #ReadParameterID_R := #Inputdata_RW_Drv2PLC.ReadParameterID_R;
   #WriteParameterID_R := #Inputdata_RW_Drv2PLC.WriteParameterID_R;
END_REGION

REGION Network 2
   RUNG wire#powerrail
      Move(in := #ReadParameterID, out1 => #Outputdata_RW_PLC2Drv.ReadParameterID)
      Move(in := #WriteParameterID, out1 => #Outputdata_RW_PLC2Drv.WriteParameterID)
      Move(in := #WriteData, out1 => #Outputdata_RW_PLC2Drv.WriteData)
   END_RUNG
   // the same network as SCL:
   #Outputdata_RW_PLC2Drv.ReadParameterID := #ReadParameterID;
   #Outputdata_RW_PLC2Drv.WriteParameterID := #WriteParameterID;
   #Outputdata_RW_PLC2Drv.WriteData := #WriteData;
END_REGION

REGION Network 3
   RUNG wire#powerrail
      Contact( #"WR-REQ" )
      Coil( #Outputdata_RW_PLC2Drv.WriteRequest."WR-REQ" )
   END_RUNG
   // the same network as SCL:
   #Outputdata_RW_PLC2Drv.WriteRequest."WR-REQ" := #"WR-REQ";
END_REGION

REGION Network 4
   RUNG wire#powerrail
      Contact( #Inputdata_RW_Drv2PLC.Read_WriteStatus."RD-ERR" )
      Coil( #"RD-ERR" )
   END_RUNG
   RUNG wire#powerrail
      Contact( #Inputdata_RW_Drv2PLC.Read_WriteStatus."SYS-BSY" )
      Coil( #"SYS-BSY" )
   END_RUNG
   RUNG wire#powerrail
      Contact( #Inputdata_RW_Drv2PLC.Read_WriteStatus."WR-END" )
      Coil( #"WR-END" )
   END_RUNG
   RUNG wire#powerrail
      Contact( #Inputdata_RW_Drv2PLC.Read_WriteStatus."WR-ERR" )
      Coil( #"WR-ERR" )
   END_RUNG
   RUNG wire#powerrail
      Contact( #Inputdata_RW_Drv2PLC.Read_WriteStatus."WR-EXE-ERR" )
      Coil( #"WR-EXE-ERR" )
   END_RUNG
   RUNG wire#powerrail
      Contact( #Inputdata_RW_Drv2PLC.Read_WriteStatus."WR-IF-ERR" )
      Coil( #"WR-IF-ERR" )
   END_RUNG
   RUNG wire#powerrail
      Contact( #Inputdata_RW_Drv2PLC.Read_WriteStatus."WR-NV-ERR" )
      Coil( #"WR-NV-ERR" )
   END_RUNG
   RUNG wire#powerrail
      Contact( #Inputdata_RW_Drv2PLC.Read_WriteStatus."WR-SET-ERR" )
      Coil( #"WR-SET-ERR" )
   END_RUNG
   // the same network as SCL:
   #"RD-ERR" := #Inputdata_RW_Drv2PLC.Read_WriteStatus."RD-ERR";
   #"SYS-BSY" := #Inputdata_RW_Drv2PLC.Read_WriteStatus."SYS-BSY";
   #"WR-END" := #Inputdata_RW_Drv2PLC.Read_WriteStatus."WR-END";
   #"WR-ERR" := #Inputdata_RW_Drv2PLC.Read_WriteStatus."WR-ERR";
   #"WR-EXE-ERR" := #Inputdata_RW_Drv2PLC.Read_WriteStatus."WR-EXE-ERR";
   #"WR-IF-ERR" := #Inputdata_RW_Drv2PLC.Read_WriteStatus."WR-IF-ERR";
   #"WR-NV-ERR" := #Inputdata_RW_Drv2PLC.Read_WriteStatus."WR-NV-ERR";
   #"WR-SET-ERR" := #Inputdata_RW_Drv2PLC.Read_WriteStatus."WR-SET-ERR";
END_REGION
END_FUNCTION_BLOCK

FUNCTION_BLOCK "POS3_0_Melden_Visu"
{ S7_Optimized_Access := 'TRUE' }
VERSION : 0.1
   VAR 
      "Taktzeitermittlung_mit_WT-Wechsel" : "Taktzeitermittlung_Start_Stop_V1_0";
      Taktzeitermittlung : "Taktzeitermittlung_Start_Stop_V1_0";
      R_TRIG_Init_Achse_1 {InstructionName := 'R_TRIG'; LibVersion := '1.0'} : R_TRIG;
      R_TRIG_Init_Achse_1_Positionen {InstructionName := 'R_TRIG'; LibVersion := '1.0'} : R_TRIG;
      R_TRIG_Init_Achse_2 {InstructionName := 'R_TRIG'; LibVersion := '1.0'} : R_TRIG;
      R_TRIG_Init_Achse_2_Positionen {InstructionName := 'R_TRIG'; LibVersion := '1.0'} : R_TRIG;
      Zyklen_für_Durchschnittszeit { ExternalAccessible := 'False'; ExternalVisible := 'False'; ExternalWritable := 'False'} : Int;
      Summe { ExternalAccessible := 'False'; ExternalVisible := 'False'; ExternalWritable := 'False'} : Real;
   END_VAR

   VAR_TEMP 
      Manuell_Zylinder_1 : Int;   // manuelle Ansteuerung Pneumatik
      Manuell_Zylinder_2 : Int;
      Manuell_Zylinder_3 : Int;
      Manuell_Zylinder_4 : Int;
      Manuell_Einzellschritt_1 : Int;
      Manuell_Einzellschritt_2 : Int;
      Manuell_Einzellschritt_3 : Int;
      Manuell_Einzellschritt_4 : Int;
      Manuell_Achse_1 : Int;   // manuelle Ansteuerung Achse 1 Seite1
      Manuell_Positionen_1_Achse_1 : Int;   // manuelle Ansteuerung Achse 1 Seite 2
      Manuell_Positionen_2_Achse_1 : Int;
      Manuell_Positionen_3_Achse_1 : Int;
      Manuell_Achse_2 : Int;
      Manuell_Positionen_1_Achse_2 : Int;
      Manuell_Positionen_2_Achse_2 : Int;
      Manuell_Positionen_3_Achse_2 : Int;
      Manuell_Achse_3 : Int;
      Manuell_Positionen_1_Achse_3 : Int;
      Manuell_Positionen_2_Achse_3 : Int;
      Manuell_Positionen_3_Achse_3 : Int;
      Manuell_Achse_4 : Int;
      Manuell_Positionen_1_Achse_4 : Int;
      Manuell_Positionen_2_Achse_4 : Int;
      Manuell_Positionen_3_Achse_4 : Int;
      i : Int;
      j : Int;
      "Manuell_P-Preset_1_Achse_1" : Int;   // manuelle Ansteuerung Achse 1 Seite 2
      "Manuell_P-Preset_1_Achse_2" : Int;   // manuelle Ansteuerung Achse 1 Seite 2
   END_VAR


BEGIN
	REGION Taktzeit  
	    
	    #Taktzeitermittlung(E_Starttrigger:="POS3_0_Signal".Station.SK_Aktiv,
	                    A_letzteZykluszeit=>"HMI_Statistik"."Letzte Zykluszeit_POS_3_0",
	                    A_letze10Zyklen=>"POS3_0_Signal".Taktzeit);
	
	"HMI_Statistik"."Letzte Zykluszeit_POS_3_0_in_s" := TIME_TO_DINT("HMI_Statistik"."Letzte Zykluszeit_POS_3_0") / 1000.0;
	
	#i := 0;
	FOR #i := 0 TO 10 DO
	    "HMI_Statistik".Zykluszeit_POS_3_0_in_s[#i] := TIME_TO_DINT("POS3_0_Signal".Taktzeit[#i]) / 1000.0;
	END_FOR;
	
	// Durchschnitt der aktuellen Istzyklen aber maximal 10 Zykluszeiten
	#Summe := 0.0;
	
	IF "POS3_0_Signal".Istzyklen < 10 THEN
	    #Zyklen_für_Durchschnittszeit := "POS3_0_Signal".Istzyklen;
	ELSE
	    #Zyklen_für_Durchschnittszeit := 10;
	END_IF;
	
	FOR #i := 1 TO #Zyklen_für_Durchschnittszeit DO
	    #Summe := #Summe + "HMI_Statistik".Zykluszeit_POS_3_0_in_s[#i];
	END_FOR;
	
	IF "POS3_0_Signal".Istzyklen <= 0 THEN
	    "HMI_Statistik"."Durchschnitt Zykluszeit_POS_3_0" := 0.0;
	ELSE
	    "HMI_Statistik"."Durchschnitt Zykluszeit_POS_3_0" := #Summe / #Zyklen_für_Durchschnittszeit;
	END_IF;
	
	// Restlaufzeit
	"POS3_0_Signal".Restzyklen := "POS3_0_Signal".Sollzyklen - "POS3_0_Signal".Istzyklen;
	
	"HMI_Statistik".Restlaufzeit_POS_3_0 := "POS3_0_Signal".Restzyklen * "HMI_Statistik"."Durchschnitt Zykluszeit_POS_3_0";
	
	
	END_REGION
	
	REGION Visu
	    
	    //Bildnummern
	    #Manuell_Zylinder_1 := 3300;
	    #Manuell_Zylinder_2 := 3301;
	    // #Manuell_Zylinder_3 := ;
	    // #Manuell_Zylinder_4:=  ;
	    // #Manuell_Einzellschritt_1:=  ;
	    // #Manuell_Einzellschritt_2:=  ;
	    // #Manuell_Einzellschritt_3:=  ;
	    // #Manuell_Einzellschritt_4:=  ;
	    #Manuell_Achse_1 := 3400;
	    #Manuell_Positionen_1_Achse_1 :=3401;
	    #"Manuell_P-Preset_1_Achse_1" := 3404;
	    // #Manuell_Positionen_2_Achse_1:= ;
	    // #Manuell_Positionen_3_Achse_1:= ;
	     #Manuell_Achse_2 := 3402;
	     #Manuell_Positionen_1_Achse_2 := 3403;
	     #"Manuell_P-Preset_1_Achse_2" := 3405;
	    // #Manuell_Positionen_2_Achse_2:=  ;
	    // #Manuell_Positionen_3_Achse_2:=  ;
	    // #Manuell_Achse_3:=  ;
	    // #Manuell_Positionen_1_Achse_3:=  ;
	    // #Manuell_Positionen_2_Achse_3:=  ;
	    // #Manuell_Positionen_3_Achse_3:=  ;
	    // #Manuell_Achse_4:=  ;
	    // #Manuell_Positionen_1_Achse_4:=  ;
	    // #Manuell_Positionen_2_Achse_4:=  ;
	    // #Manuell_Positionen_3_Achse_4:=  ;
	    // 
	    
	    
	    REGION Wartezeit Ist gesteckt
	        "POS3_0_Signal"."Wartezeit Ist gesteckt" := TIME_TO_DINT("POS3_0_SK_Ablauf_DB"."Wartezeit - Messmethode_AUS".T) / 1000.0;
	      
	    END_REGION
	    
	END_REGION
	
	
	
	REGION Allgemein
	    //Allgemein 
	    
	    "HMI_BETR_ART_POS".POS3_0.Status_Sicher := FALSE;
	    "HMI_BETR_ART_POS".POS3_0.Status_Anwahl := "POS3_0_Signal".Schrittkette.TAP_ON;
	    "HMI_BETR_ART_POS".POS3_0.SNr := "POS3_0_Signal".Schrittkette.S_NO;
	    
	    // Status Richten
	    IF "POS3_0_Signal".Station.SK_Richten_gestartet THEN
	        "HMI_BETR_ART_POS".POS3_0.Status_Richten := 1;
	    ELSIF "Global_Signal"."M_Grundstellung_POS3.0" THEN
	        "HMI_BETR_ART_POS".POS3_0.Status_Richten := 2;
	    ELSE
	        "HMI_BETR_ART_POS".POS3_0.Status_Richten := 0;
	    END_IF;
	   
	    
	    // Status Schrittkette
	    IF "POS3_0_Signal".Station.SK_Aktiv AND NOT "POS3_0_Signal".Station.SK_Fertig THEN
	        "HMI_BETR_ART_POS".POS3_0.Status_Schrittkette := 1;    //  1 = Schrittkette läuft
	    ELSIF "POS3_0_Signal".Station.SK_Fertig THEN
	        "HMI_BETR_ART_POS".POS3_0.Status_Schrittkette := 2;    //  2 = Schrittkette fertig
	    ELSIF "POS3_0_Signal".Schrittkette.ERR_FLT  THEN
	        "HMI_BETR_ART_POS".POS3_0.Status_Schrittkette := 3;    //  3 = Taktzeit max Störung
	    ELSE
	        "HMI_BETR_ART_POS".POS3_0.Status_Schrittkette := 0;    //  0 = Schrittkette AUS    
	    END_IF;
	   
	END_REGION
	
	REGION Manuell
	    // Manuellaufruf der Station über Bildanwahl
	     REGION Zylinder_1
	         IF ("HMI_SYS"."Aktueller Bildschirm" = #Manuell_Zylinder_1) THEN
	            
	             "HMI_COM".Manuell_Zylinder1."0_Aus_1_Ventil_2_Antrieb_3_Signal" := 3;
	             IF "DE_POS3_0_Endlage_Überlastzylinder" THEN
	                 "HMI_COM".Manuell_Zylinder1.Status := 0;
	             ELSE
	                 "HMI_COM".Manuell_Zylinder1.Status := 1;
	             END_IF;
	            
	            
	             "HMI_COM".Manuell_Zylinder2."0_Aus_1_Ventil_2_Antrieb_3_Signal" := 3;
	             IF FALSE THEN
	                 "HMI_COM".Manuell_Zylinder2.Status := 1;
	             ELSE
	                 "HMI_COM".Manuell_Zylinder2.Status := 0;
	             END_IF;
	            
	                
	             "HMI_COM".Manuell_Zylinder3."0_Aus_1_Ventil_2_Antrieb_3_Signal" := 3;
	             IF false THEN
	                 "HMI_COM".Manuell_Zylinder3.Status := 1;
	             ELSE
	                 "HMI_COM".Manuell_Zylinder3.Status := 0;
	             END_IF;
	            
	             
	              "HMI_COM".Manuell_Zylinder4."0_Aus_1_Ventil_2_Antrieb_3_Signal" := 3;
	              IF FALSE THEN
	                  "HMI_COM".Manuell_Zylinder4.Status := 1;
	              ELSE
	                  "HMI_COM".Manuell_Zylinder4.Status := 0;
	              END_IF;
	             
	             
	            
	            
	        //     // //Manuelle Ansteuerung Zylinder
	        //      // := "HMI_COM".Manuell_Zylinder1.GS;
	        //      // := "HMI_COM".Manuell_Zylinder1.AS1;
	        
	        //      // := "HMI_COM".Manuell_Zylinder2.GS;
	        //      // := "HMI_COM".Manuell_Zylinder2.AS1;
	            
	        //      // := "HMI_COM".Manuell_Zylinder3.GS;
	        //      // := "HMI_COM".Manuell_Zylinder3.AS1;
	            
	        //      // := "HMI_COM".Manuell_Zylinder4.GS;
	        //      // := "HMI_COM".Manuell_Zylinder4.AS1;
	            
	        //     "HMI_COM".Manuell_Zylinder1.GS := false;
	        //     "HMI_COM".Manuell_Zylinder1.AS1 := false;
	        //     "HMI_COM".Manuell_Zylinder2.GS := false;
	        //     "HMI_COM".Manuell_Zylinder2.AS1 := false;
	        //     "HMI_COM".Manuell_Zylinder3.GS := false;
	        //     "HMI_COM".Manuell_Zylinder3.AS1 := false;
	        //     "HMI_COM".Manuell_Zylinder4.GS := false;
	        //     "HMI_COM".Manuell_Zylinder4.AS1 := false;
	            
	            
	        //     //Rückmeldung Ansteuerung aktiv
	        //     "HMI_COM".Manuell_Zylinder1.DA_GS := FALSE;
	        //     "HMI_COM".Manuell_Zylinder1.DA_AS1 := FALSE;
	        //     "HMI_COM".Manuell_Zylinder1.DA_AS2 := FALSE;
	            
	        //     "HMI_COM".Manuell_Zylinder2.DA_GS := FALSE;
	        //     "HMI_COM".Manuell_Zylinder2.DA_AS1 := FALSE;
	        //     "HMI_COM".Manuell_Zylinder2.DA_AS2 := FALSE;
	            
	        //     "HMI_COM".Manuell_Zylinder3.DA_GS := FALSE;
	        //     "HMI_COM".Manuell_Zylinder3.DA_AS1 := FALSE;
	        //     "HMI_COM".Manuell_Zylinder3.DA_AS2 := FALSE;
	            
	        //     "HMI_COM".Manuell_Zylinder4.DA_GS := FALSE;
	        //     "HMI_COM".Manuell_Zylinder4.DA_AS1 := FALSE;
	        //     "HMI_COM".Manuell_Zylinder4.DA_AS2 := FALSE;
	            
	         END_IF;
	     END_REGION ;
	  
	 
	 
	    
	    REGION Antrieb 1 Positionierachse
	        // Initialisieren der Steuerwerte 
	        #R_TRIG_Init_Achse_1(CLK := "HMI_SYS"."Aktueller Bildschirm" = #Manuell_Achse_1);
	        IF #R_TRIG_Init_Achse_1.Q THEN
	            "HMI_COM".HMI_Achse_Steuerung.E_Sollwert_Manuell := "POS3_0_Signal"."-1001T1 Oriental_Steuerung".E_DDO_Pos;
	            "HMI_COM".HMI_Achse_Steuerung.E_Verfahrweg := "POS3_0_Signal"."-1001T1 Oriental_Steuerung".E_Schrittweite;
	            "HMI_COM".HMI_Achse_Steuerung.E_Geschwindigkeit_manuell_in_Prozent := "POS3_0_Signal"."-1001T1 Oriental_Steuerung".E_DDO_Vel;
	        END_IF;
	        
	        
	        IF ("HMI_SYS"."Aktueller Bildschirm" = #Manuell_Achse_1) THEN
	            "POS3_0_Signal"."-1001T1 Oriental_Steuerung".E_ZHOME := "HMI_COM".HMI_Achse_Steuerung.E_Start_Referenzieren;
	            "HMI_COM".HMI_Achse_Steuerung.A_StatusWord := "POS3_0_Signal"."-1001T1 Oriental_Steuerung".A_StatusWord;
	            "HMI_COM".HMI_Achse_Steuerung.E_Drehachse := false;
	            "HMI_COM".HMI_Achse_Steuerung.E_Achstyp := 3;
	            
	            "HMI_COM".HMI_Achse_Steuerung.A_Istwert := REAL_TO_LREAL("POS3_0_Signal"."-1001T1 Oriental_Steuerung".A_FBposition);
	            "HMI_COM".HMI_Achse_Steuerung.A_Softw_ES_min := "POS3_0_Signal"."-1001T1 Oriental_Positionen".A_Softw_ES_min_mm;
	            "HMI_COM".HMI_Achse_Steuerung.A_Softw_ES_max := "POS3_0_Signal"."-1001T1 Oriental_Positionen".A_Softw_ES_max_mm;
	            
	            "POS3_0_Signal"."-1001T1 Oriental_Steuerung".E_DDO_Pos := LREAL_TO_REAL("HMI_COM".HMI_Achse_Steuerung.E_Sollwert_Manuell);
	            "POS3_0_Signal"."-1001T1 Oriental_Steuerung".E_Schrittweite := LREAL_TO_REAL("HMI_COM".HMI_Achse_Steuerung.E_Verfahrweg);
	            "POS3_0_Signal"."-1001T1 Oriental_Steuerung".E_DDO_Vel := LREAL_TO_REAL("HMI_COM".HMI_Achse_Steuerung.E_Geschwindigkeit_manuell_in_Prozent);
	            "POS3_0_Signal"."-1001T1 Oriental_Steuerung".E_DDO_Acc := 100.0;
	            "POS3_0_Signal"."-1001T1 Oriental_Steuerung".E_DDO_Dec := 100.0;
	            "POS3_0_Signal"."-1001T1 Oriental_Steuerung".E_DDO_Crnt := 100;
	            
	            "POS3_0_Signal"."-1001T1 Oriental_Steuerung".E_Schrittweite_pos := "HMI_COM".HMI_Achse_Steuerung.E_Tipp_pos;
	            "POS3_0_Signal"."-1001T1 Oriental_Steuerung".E_Schrittweite_neg := "HMI_COM".HMI_Achse_Steuerung.E_Tipp_neg;
	            "POS3_0_Signal"."-1001T1 Oriental_Steuerung".E_Trig_Manuell := "HMI_COM".HMI_Achse_Steuerung.E_Start_manuell;
	            "POS3_0_Signal"."-1001T1 Oriental_Steuerung"."E_FW-JOG" := "HMI_COM".HMI_Achse_Steuerung.E_jog_pos;
	            "POS3_0_Signal"."-1001T1 Oriental_Steuerung"."E_RV-JOG" := "HMI_COM".HMI_Achse_Steuerung.E_jog_neg;
	        END_IF;
	            
	            // Initialisieren der Steuerwerte 
	            #R_TRIG_Init_Achse_1_Positionen(CLK := "HMI_SYS"."Aktueller Bildschirm" = #Manuell_Positionen_1_Achse_1);
	        IF #R_TRIG_Init_Achse_1_Positionen.Q THEN
	                "HMI_COM".HMI_Achse_POS_Überschreiben.Wert_Position_Überschreiben[0] := "POS3_0_Signal"."-1001T1 Oriental_Positionen".Soll_Position[0];
	                "HMI_COM".HMI_Achse_POS_Überschreiben.Wert_Speed_Überschreiben[0] := "POS3_0_Signal"."-1001T1 Oriental_Positionen".Geschwindigkeit[0];
	                 
	                "HMI_COM".HMI_Achse_POS_Überschreiben.Wert_Position_Überschreiben[1] := "POS3_0_Signal"."-1001T1 Oriental_Positionen".Soll_Position[1];
	                "HMI_COM".HMI_Achse_POS_Überschreiben.Wert_Speed_Überschreiben[1] := "POS3_0_Signal"."-1001T1 Oriental_Positionen".Geschwindigkeit[1];
	                
	                "HMI_COM".HMI_Achse_POS_Überschreiben.Wert_Position_Überschreiben[2] := "POS3_0_Signal"."-1001T1 Oriental_Positionen".Soll_Position[2];
	                "HMI_COM".HMI_Achse_POS_Überschreiben.Wert_Speed_Überschreiben[2] := "POS3_0_Signal"."-1001T1 Oriental_Positionen".Geschwindigkeit[2];
	                
	                "HMI_COM".HMI_Achse_POS_Überschreiben.Wert_Position_Überschreiben[3] := "POS3_0_Signal"."-1001T1 Oriental_Positionen".Soll_Position[3];
	                "HMI_COM".HMI_Achse_POS_Überschreiben.Wert_Speed_Überschreiben[3] := "POS3_0_Signal"."-1001T1 Oriental_Positionen".Geschwindigkeit[3];
	                
	                "HMI_COM".HMI_Achse_POS_Überschreiben.Wert_Position_Überschreiben[4] := "POS3_0_Signal"."-1001T1 Oriental_Positionen".Soll_Position[4];
	                "HMI_COM".HMI_Achse_POS_Überschreiben.Wert_Speed_Überschreiben[4] := "POS3_0_Signal"."-1001T1 Oriental_Positionen".Geschwindigkeit[4];
	                
	                "HMI_COM".HMI_Achse_POS_Überschreiben.Wert_Position_Überschreiben[5] := "POS3_0_Signal"."-1001T1 Oriental_Positionen".Soll_Position[5];
	                "HMI_COM".HMI_Achse_POS_Überschreiben.Wert_Speed_Überschreiben[5] := "POS3_0_Signal"."-1001T1 Oriental_Positionen".Geschwindigkeit[5];
	                
	        END_IF;
	            
	            
	        IF ("HMI_SYS"."Aktueller Bildschirm" = #Manuell_Positionen_1_Achse_1) THEN
	                
	            
	            "HMI_COM".HMI_Achse_Steuerung.A_StatusWord := "POS3_0_Signal"."-1001T1 Oriental_Steuerung".A_StatusWord;
	            "HMI_COM".HMI_Achse_Steuerung.E_Drehachse := false;
	            "HMI_COM".HMI_Achse_Steuerung.A_Istwert := REAL_TO_LREAL("POS3_0_Signal"."-1001T1 Oriental_Steuerung".A_FBposition);
	            "HMI_COM".HMI_Achse_Steuerung.A_Softw_ES_min := "POS3_0_Signal"."-1001T1 Oriental_Positionen".A_Softw_ES_min_mm;
	            "HMI_COM".HMI_Achse_Steuerung.A_Softw_ES_max := "POS3_0_Signal"."-1001T1 Oriental_Positionen".A_Softw_ES_max_mm;
	            
	            
	            "HMI_COM".HMI_Achse_Position.Soll_Wert_in_mm_Position[0] := "POS3_0_Signal"."-1001T1 Oriental_Positionen".Soll_Position[0];
	            "HMI_COM".HMI_Achse_Position.Soll_Wert_in_mm_Position[1] := "POS3_0_Signal"."-1001T1 Oriental_Positionen".Soll_Position[1];
	            "HMI_COM".HMI_Achse_Position.Soll_Wert_in_mm_Position[2] := "POS3_0_Signal"."-1001T1 Oriental_Positionen".Soll_Position[2];
	            "HMI_COM".HMI_Achse_Position.Soll_Wert_in_mm_Position[3] := "POS3_0_Signal"."-1001T1 Oriental_Positionen".Soll_Position[3];
	            "HMI_COM".HMI_Achse_Position.Soll_Wert_in_mm_Position[4] := "POS3_0_Signal"."-1001T1 Oriental_Positionen".Soll_Position[4];
	            "HMI_COM".HMI_Achse_Position.Soll_Wert_in_mm_Position[5] := "POS3_0_Signal"."-1001T1 Oriental_Positionen".Soll_Position[5];
	            
	            "HMI_COM".HMI_Achse_Position.POS_OK_Position[0] := "POS3_0_Signal"."-1001T1 Oriental_Positionen".POS_OK_Position[0];
	            "HMI_COM".HMI_Achse_Position.POS_OK_Position[1] := "POS3_0_Signal"."-1001T1 Oriental_Positionen".POS_OK_Position[1];
	            "HMI_COM".HMI_Achse_Position.POS_OK_Position[2] := "POS3_0_Signal"."-1001T1 Oriental_Positionen".POS_OK_Position[2];
	            "HMI_COM".HMI_Achse_Position.POS_OK_Position[3] := "POS3_0_Signal"."-1001T1 Oriental_Positionen".POS_OK_Position[3];
	            "HMI_COM".HMI_Achse_Position.POS_OK_Position[4] := "POS3_0_Signal"."-1001T1 Oriental_Positionen".POS_OK_Position[4];
	            "HMI_COM".HMI_Achse_Position.POS_OK_Position[5] := "POS3_0_Signal"."-1001T1 Oriental_Positionen".POS_OK_Position[5];
	            
	            "HMI_COM".HMI_Achse_Position.Soll_Speed_in_Prozent_Position[0] := "POS3_0_Signal"."-1001T1 Oriental_Positionen".Geschwindigkeit[0];
	            "HMI_COM".HMI_Achse_Position.Soll_Speed_in_Prozent_Position[1] := "POS3_0_Signal"."-1001T1 Oriental_Positionen".Geschwindigkeit[1];
	            "HMI_COM".HMI_Achse_Position.Soll_Speed_in_Prozent_Position[2] := "POS3_0_Signal"."-1001T1 Oriental_Positionen".Geschwindigkeit[2];
	            "HMI_COM".HMI_Achse_Position.Soll_Speed_in_Prozent_Position[3] := "POS3_0_Signal"."-1001T1 Oriental_Positionen".Geschwindigkeit[3];
	            "HMI_COM".HMI_Achse_Position.Soll_Speed_in_Prozent_Position[4] := "POS3_0_Signal"."-1001T1 Oriental_Positionen".Geschwindigkeit[4];
	            "HMI_COM".HMI_Achse_Position.Soll_Speed_in_Prozent_Position[5] := "POS3_0_Signal"."-1001T1 Oriental_Positionen".Geschwindigkeit[5];
	            
	            "POS3_0_Signal"."-1001T1 Oriental_Positionen".Start_POS_Position[0] := "HMI_COM".HMI_Achse_Position.Start_POS_Position[0];
	            "POS3_0_Signal"."-1001T1 Oriental_Positionen".Start_POS_Position[1] := "HMI_COM".HMI_Achse_Position.Start_POS_Position[1];
	            "POS3_0_Signal"."-1001T1 Oriental_Positionen".Start_POS_Position[2] := "HMI_COM".HMI_Achse_Position.Start_POS_Position[2];
	            "POS3_0_Signal"."-1001T1 Oriental_Positionen".Start_POS_Position[3] := "HMI_COM".HMI_Achse_Position.Start_POS_Position[3];
	            "POS3_0_Signal"."-1001T1 Oriental_Positionen".Start_POS_Position[4] := "HMI_COM".HMI_Achse_Position.Start_POS_Position[4];
	            "POS3_0_Signal"."-1001T1 Oriental_Positionen".Start_POS_Position[5] := "HMI_COM".HMI_Achse_Position.Start_POS_Position[5];
	            
	            
	            IF "HMI_COM".HMI_Achse_POS_Überschreiben.Trig_Position_Überschreiben[0] THEN
	                "POS3_0_Signal"."-1001T1 Oriental_Positionen".Soll_Position[0] := "HMI_COM".HMI_Achse_POS_Überschreiben.Wert_Position_Überschreiben[0];
	                "POS3_0_Signal"."-1001T1 Oriental_Positionen".Geschwindigkeit[0]:= "HMI_COM".HMI_Achse_POS_Überschreiben.Wert_Speed_Überschreiben[0];
	            END_IF;
	            
	            IF "HMI_COM".HMI_Achse_POS_Überschreiben.Trig_Position_Überschreiben[1] THEN
	                "POS3_0_Signal"."-1001T1 Oriental_Positionen".Soll_Position[1] := "HMI_COM".HMI_Achse_POS_Überschreiben.Wert_Position_Überschreiben[1];
	                "POS3_0_Signal"."-1001T1 Oriental_Positionen".Geschwindigkeit[1] := "HMI_COM".HMI_Achse_POS_Überschreiben.Wert_Speed_Überschreiben[1];
	            END_IF;
	            
	            IF "HMI_COM".HMI_Achse_POS_Überschreiben.Trig_Position_Überschreiben[2] THEN
	                "POS3_0_Signal"."-1001T1 Oriental_Positionen".Soll_Position[2] := "HMI_COM".HMI_Achse_POS_Überschreiben.Wert_Position_Überschreiben[2];
	                "POS3_0_Signal"."-1001T1 Oriental_Positionen".Geschwindigkeit[2] := "HMI_COM".HMI_Achse_POS_Überschreiben.Wert_Speed_Überschreiben[2];
	            END_IF;
	            
	            IF "HMI_COM".HMI_Achse_POS_Überschreiben.Trig_Position_Überschreiben[3] THEN
	                "POS3_0_Signal"."-1001T1 Oriental_Positionen".Soll_Position[3] := "HMI_COM".HMI_Achse_POS_Überschreiben.Wert_Position_Überschreiben[3];
	                "POS3_0_Signal"."-1001T1 Oriental_Positionen".Geschwindigkeit[3] := "HMI_COM".HMI_Achse_POS_Überschreiben.Wert_Speed_Überschreiben[3];
	            END_IF;
	            
	            IF "HMI_COM".HMI_Achse_POS_Überschreiben.Trig_Position_Überschreiben[4] THEN
	                "POS3_0_Signal"."-1001T1 Oriental_Positionen".Soll_Position[4] := "HMI_COM".HMI_Achse_POS_Überschreiben.Wert_Position_Überschreiben[4];
	                "POS3_0_Signal"."-1001T1 Oriental_Positionen".Geschwindigkeit[4] := "HMI_COM".HMI_Achse_POS_Überschreiben.Wert_Speed_Überschreiben[4];
	            END_IF;
	            
	            IF "HMI_COM".HMI_Achse_POS_Überschreiben.Trig_Position_Überschreiben[5] THEN
	                "POS3_0_Signal"."-1001T1 Oriental_Positionen".Soll_Position[5] := "HMI_COM".HMI_Achse_POS_Überschreiben.Wert_Position_Überschreiben[5];
	                "POS3_0_Signal"."-1001T1 Oriental_Positionen".Geschwindigkeit[5] := "HMI_COM".HMI_Achse_POS_Überschreiben.Wert_Speed_Überschreiben[5];
	            END_IF;
	            
	            
	            
	        END_IF;
	        
	        
	        IF ("HMI_SYS"."Aktueller Bildschirm" = #"Manuell_P-Preset_1_Achse_1") THEN
	            "HMI_COM".HMI_Achse_Steuerung.A_StatusWord := "POS3_0_Signal"."-1001T1 Oriental_Steuerung".A_StatusWord;
	            "HMI_COM".HMI_Achse_Steuerung.E_Drehachse := false;
	            "HMI_COM".HMI_Achse_Steuerung.A_Istwert := REAL_TO_LREAL("POS3_0_Signal"."-1001T1 Oriental_Steuerung".A_FBposition);
	        END_IF;
	        
	    END_REGION
	    
	    
	    
	    REGION Antrieb 2 Drehachse
	        // Initialisieren der Steuerwerte 
	        #R_TRIG_Init_Achse_2(CLK := "HMI_SYS"."Aktueller Bildschirm" = #Manuell_Achse_2);
	        IF #R_TRIG_Init_Achse_2.Q THEN
	            "HMI_COM".HMI_Achse_Steuerung.E_Sollwert_Manuell := "POS3_0_Signal"."-1002T1 Oriental_Steuerung".E_DDO_Pos;
	            "HMI_COM".HMI_Achse_Steuerung.E_Verfahrweg := "POS3_0_Signal"."-1002T1 Oriental_Steuerung".E_Schrittweite;
	            "HMI_COM".HMI_Achse_Steuerung.E_Geschwindigkeit_manuell_in_Prozent := "POS3_0_Signal"."-1002T1 Oriental_Steuerung".E_DDO_Vel;
	        END_IF;
	        
	        
	        IF ("HMI_SYS"."Aktueller Bildschirm" = #Manuell_Achse_2) THEN
	            "POS3_0_Signal"."-1002T1 Oriental_Steuerung".E_ZHOME := "HMI_COM".HMI_Achse_Steuerung.E_Start_Referenzieren;
	            "HMI_COM".HMI_Achse_Steuerung.A_StatusWord := "POS3_0_Signal"."-1001T1 Oriental_Steuerung".A_StatusWord;
	            "HMI_COM".HMI_Achse_Steuerung.E_Drehachse := true;
	            "HMI_COM".HMI_Achse_Steuerung.E_Achstyp := 3;
	            
	            "HMI_COM".HMI_Achse_Steuerung.A_Istwert := REAL_TO_LREAL("POS3_0_Signal"."-1002T1 Oriental_Steuerung".A_FBposition);
	            "HMI_COM".HMI_Achse_Steuerung.A_Softw_ES_min := "POS3_0_Signal"."-1002T1 Oriental_Positionen".A_Softw_ES_min_mm;
	            "HMI_COM".HMI_Achse_Steuerung.A_Softw_ES_max := "POS3_0_Signal"."-1002T1 Oriental_Positionen".A_Softw_ES_max_mm;
	            
